Omron Sysmac Studio project TP - Automaçao (Sysmac Studio 1.56.0.64011, StandardProject)

# Controller new_Controller_0: NX1P2-9B24DT1 version 1.42
Task PrimaryTask (priority 4, period or condition 4000): Program0
Library OEN_Communication_V1_0_22 1.0.22 (contents left out)

VAR_GLOBAL
    Trama : ARRAY[0..3] OF OEN\Modbus\sModbusReq := [(Enable := True, NodeAdr := 1, FunctionCode := Fn02_ReadDiscreteInputs, Read := (StartAddressRemote := 0, StartAddressLocal := 0, Count := 49), Write := (StartAddressRemote := 0, StartAddressLocal := 0, Count := 0)), (Enable := True, NodeAdr := 1, FunctionCode := Fn15_WriteMultipleCoils, Read := (StartAddressRemote := 0, StartAddressLocal := 0, Count := 0), Write := (StartAddressRemote := 0, StartAddressLocal := 0, Count := 129)), (Enable := True, NodeAdr := 1, FunctionCode := Fn04_ReadInputRegisters, Read := (StartAddressRemote := 0, StartAddressLocal := 0, Count := 10), Write := (StartAddressRemote := 0, StartAddressLocal := 0, Count := 0)), (Enable := True, NodeAdr := 1, FunctionCode := Fn16_WriteMultipleRegisters, Read := (StartAddressRemote := 0, StartAddressLocal := 0, Count := 0), Write := (StartAddressRemote := 0, StartAddressLocal := 0, Count := 10))];  (* Trama *)
    out_Dig : ARRAY[0..130] OF BOOL;  (* Saidas digitais *)
    in_Dig : ARRAY[0..50] OF BOOL;  (* Entradas digitais *)
    in_Analog : ARRAY[0..10] OF WORD;  (* Entradas analogicas *)
    out_Analog : ARRAY[0..10] OF WORD;  (* Saidas analogicas *)
    BIO_Input_Bit_00 : BOOL;  (* Botão fisico; at BuiltInIO://cpu/#0/Input_Bit_00 *)
    BIO_Output_Bit_00 : BOOL;  (* Led Verde - Fisico; at BuiltInIO://cpu/#0/Output_Bit_00 *)
    BIO_Output_Bit_01 : BOOL;  (* Led Amarelo - Fisico; at BuiltInIO://cpu/#0/Output_Bit_01 *)
    BIO_Output_Bit_02 : BOOL;  (* Led Vermelho - Fisico; at BuiltInIO://cpu/#0/Output_Bit_02 *)
    ANALOG_Ch1_Analog_Output_Value : INT;  (* at BuiltInIO://opt/#0/Ch1_Analog_Output_Value *)
    Encomenda_Azul : DINT;  (* Numero de peça desta cor por encomenda *)
    Encomenda_Verde : DINT;  (* Numero de peça desta cor por encomenda *)
    Encomenda_Cinza : DINT;  (* Numero de peça desta cor por encomenda *)
    Peca_Boa_Azul : DINT;  (* Contador de peças boas produzidas *)
    Peca_Boa_Verde : DINT;  (* Contador de peças boas produzidas *)
    Peca_Boa_Cinza : DINT;  (* Contador de peças boas produzidas *)
    Peca_Lixo_Azul : DINT;  (* Contador de peças com defeito produzidas *)
    Peca_Lixo_Verde : DINT;  (* Contador de peças com defeito produzidas *)
    Peca_Lixo_Cinza : DINT;  (* Contador de peças com defeito produzidas *)
    Peca_Stock_Azul : DINT;  (* Contador de peças que foram para stock *)
    Peca_Stock_Verde : DINT;  (* Contador de peças que foram para stock *)
    Peca_Stock_Cinza : DINT;  (* Contador de peças que foram para stock *)
    HMI_Emitter : BOOL;
    HMI_R8 : BOOL;
    HMI_R0 : BOOL;
    HMI_R1 : BOOL;
    HMI_R3 : BOOL;
    HMI_R2 : BOOL;
    HMI_R4 : BOOL;
    HMI_R5 : BOOL;
    HMI_Alarme : BOOL;
    HMI_LG_10 : BOOL;
    HMI_LG_11 : BOOL;
    HMI_LG_12 : BOOL;
    HMI_LG_13 : BOOL;
    HMI_LG_14 : BOOL;
    HMI_LG_15 : BOOL;
    HMI_LG_18 : BOOL;
    HMI_LG_19 : BOOL;
    HMI_LY_10 : BOOL;
    HMI_LY_11 : BOOL;
    HMI_LY_12 : BOOL;
    HMI_LY_13 : BOOL;
    HMI_LY_14 : BOOL;
    HMI_LY_15 : BOOL;
    HMI_LY_18 : BOOL;
    HMI_LY_19 : BOOL;
    HMI_LR_10 : BOOL;
    HMI_LR_11 : BOOL;
    HMI_LR_12 : BOOL;
    HMI_LR_13 : BOOL;
    HMI_LR_14 : BOOL;
    HMI_LR_15 : BOOL;
    HMI_LR_18 : BOOL;
    HMI_LR_19 : BOOL;
    HMI_PP0_X : BOOL;
    HMI_PP1_X : BOOL;
    HMI_PP2_X : BOOL;
    HMI_PP0_Z : BOOL;
    HMI_PP1_Z : BOOL;
    HMI_PP2_Z : BOOL;
    HMI_PP0_Grab : BOOL;
    HMI_PP1_Grab : BOOL;
    HMI_PP2_Grab : BOOL;
    HMI_PP0_CW : BOOL;
    HMI_PP1_CW : BOOL;
    HMI_PP2_CW : BOOL;
    HMI_PP0_CCW : BOOL;
    HMI_PP1_CCW : BOOL;
    HMI_PP2_CCW : BOOL;
    HMI_DS0 : BOOL;
    HMI_DS1 : BOOL;
    HMI_DS2 : BOOL;
    HMI_DS3 : BOOL;
    HMI_DS4 : BOOL;
    HMI_DS5 : BOOL;
    HMI_DS6 : BOOL;
    HMI_DS7 : BOOL;
    HMI_DS8 : BOOL;
    HMI_DS9 : BOOL;
    HMI_DS10 : BOOL;
    HMI_DS11 : BOOL;
    HMI_DS12 : BOOL;
    HMI_DS13 : BOOL;
    HMI_DS14 : BOOL;
    HMI_DS15 : BOOL;
    HMI_DS16 : BOOL;
    HMI_DS17 : BOOL;
    HMI_DS18 : BOOL;
    HMI_DS19 : BOOL;
    HMI_DS20 : BOOL;
    HMI_DS21 : BOOL;
    HMI_DS22 : BOOL;
    HMI_DS23 : BOOL;
    HMI_DS24 : BOOL;
    HMI_DS25 : BOOL;
    HMI_DS26 : BOOL;
    HMI_DS27 : BOOL;
    HMI_DS28 : BOOL;
    HMI_T20 : BOOL;
    HMI_T21 : BOOL;
    HMI_T22 : BOOL;
    HMI_T23 : BOOL;
    HMI_T24 : BOOL;
    HMI_T25 : BOOL;
    HMI_T26 : BOOL;
    HMI_T27 : BOOL;
    HMI_T28 : BOOL;
    HMI_T29 : BOOL;
    HMI_T210 : BOOL;
    HMI_T211 : BOOL;
    HMI_T212 : BOOL;
    HMI_T213 : BOOL;
    HMI_T214 : BOOL;
    HMI_T215 : BOOL;
    HMI_T216 : BOOL;
    HMI_T217 : BOOL;
    HMI_T218 : BOOL;
    HMI_T219 : BOOL;
    HMI_T220 : BOOL;
    HMI_T221 : BOOL;
    HMI_T222 : BOOL;
    HMI_T223 : BOOL;
    HMI_T224 : BOOL;
    HMI_T225 : BOOL;
    HMI_T226 : BOOL;
    HMI_T227 : BOOL;
    HMI_T229 : BOOL;
    HMI_T230 : BOOL;
    HMI_T40 : BOOL;
    HMI_T41 : BOOL;
    HMI_T42 : BOOL;
    HMI_T43 : BOOL;
    HMI_T45 : BOOL;
    HMI_T46 : BOOL;
    HMI_T60 : BOOL;
    HMI_T61 : BOOL;
    HMI_T62 : BOOL;
    HMI_T63 : BOOL;
    HMI_T64 : BOOL;
    HMI_T65 : BOOL;
    HMI_T66 : BOOL;
    HMI_T67 : BOOL;
    HMI_T68 : BOOL;
    HMI_T69 : BOOL;
    HMI_CCW1 : BOOL;
    HMI_CCW0 : BOOL;
    HMI_CW2 : BOOL;
    HMI_CW3 : BOOL;
    HMI_CW4 : BOOL;
    HMI_CW5 : BOOL;
    HMI_CCW6 : BOOL;
    HMI_CCW7 : BOOL;
    HMI_CW8 : BOOL;
    HMI_CW9 : BOOL;
    HMI_CW10 : BOOL;
    HMI_CW11 : BOOL;
    HMI_CW12 : BOOL;
    HMI_CCW14 : BOOL;
    HMI_CW15 : BOOL;
    HMI_CW16 : BOOL;
    HMI_CW17 : BOOL;
    HMI_CW18 : BOOL;
    HMI_CCW20 : BOOL;
    HMI_CW21 : BOOL;
    HMI_PA3_Turn : BOOL;
    HMI_PA4_Turn : BOOL;
    HMI_PA3_Power : BOOL;
    HMI_PA4_Power : BOOL;
    HMI_B0_Power : BOOL;
    HMI_B1_Power : BOOL;
    HMI_B2_Power : BOOL;
    HMI_L0 : BOOL;
    HMI_L1 : BOOL;
    HMI_L2 : BOOL;
    HMI_MCS_0 : BOOL;
    HMI_MCS_1 : BOOL;
    HMI_MCS_2 : BOOL;
    Terminar_sessao : BOOL;  (* Sai do modo de manutenção da HMI *)
    HMI_Emissor : BOOL;
    HMI_Led_producao : BOOL;
    HMI_Led_Manutencao : BOOL;
    HMI_PP3_CCW : BOOL;
    HMI_PP3_CW : BOOL;
    HMI_BT_Linha_Principal : BOOL;
    HMI_BT_Linha_Azul : BOOL;
    HMI_BT_Linha_Verde : BOOL;
    HMI_BT_Linha_Cinza : BOOL;
    HMI_BT_Linha_Recolha : BOOL;
    VS : DINT;  (* Vision sensor *)
    Flag_Stop : BOOL;
    DS16 : BOOL;
    Encomenda_Total : DINT;
    DS28 : BOOL;
    BTSL_1 : BOOL;  (* Botão Seletor - posição 1 *)
    Page_Access : BOOL;
    HMI_Encomenda_Azul_Historico : ARRAY[1..10] OF REAL;
    HMI_Encomenda_Verde_Historico : ARRAY[1..10] OF REAL;
    HMI_Encomenda_Cinza_Historico : ARRAY[1..10] OF REAL;
    HMI_Historico_Index : INT := 1;
    Page_Access1 : BOOL;
    HMI_VoltaP : BOOL;
    HMI_VoltaRC : BOOL;
    HMI_Volta1 : BOOL;
    HMI_Volta2 : BOOL;
    HMI_Volta3 : BOOL;
    Encomenda_Pronta : BOOL;
    HMI_Flag_Stop : BOOL;
    HMI_VS : DINT;
    HMI_DS29 : BOOL;
    HMI_DS30 : BOOL;
    HMI_DS31 : BOOL;
    HMI_DS33 : BOOL;
    HMI_DS34 : BOOL;
    HMI_DS32 : BOOL;
    HMI_Emergencia : BOOL;
END_VAR

PROGRAM Program0
VAR
    ModBus_Client_PLC : OEN\Modbus\ModbusTCP_Client;  (* Bloco ModBus *)
    L0 : BOOL;  (* Lamina stop 0 *)
    L1 : BOOL;  (* Lamina stop 1 *)
    L2 : BOOL;  (* Lamina stop 2 *)
    Emitter : BOOL;  (* Emissor de peças *)
    R0 : BOOL;  (* Peças para o lixo *)
    R1 : BOOL;  (* Peças para o lixo *)
    R2 : BOOL;  (* Peças para stock *)
    R3 : BOOL;  (* Peças para o lixo *)
    R4 : BOOL;  (* Peças para stock *)
    R5 : BOOL;  (* Peças para stock *)
    R8 : BOOL;  (* Remove encomenda final *)
    BTSL_0 : BOOL;  (* Botão Seletor - posição 0 *)
    BTS : BOOL;  (* Botão Start *)
    BTE : BOOL;  (* Botão Emergencia *)
    BTSP : BOOL;  (* Botão Stop *)
    BTR : BOOL;  (* Botão Reset *)
    A2 : BOOL;  (* Alarme *)
    LG_10 : BOOL;  (* Led Verde - semaforo 10 *)
    LG_11 : BOOL;  (* Led Verde - semaforo 11 *)
    LG_12 : BOOL;  (* Led Verde - semaforo 12 *)
    LG_13 : BOOL;  (* Led Verde - semaforo 13 *)
    LG_14 : BOOL;  (* Led Verde - semaforo 14 *)
    LG_15 : BOOL;  (* Led Verde - semaforo 15 *)
    LG_18 : BOOL;  (* Led Verde - semaforo 18 *)
    LG_19 : BOOL;  (* Led Verde - semaforo 19 *)
    LR_10 : BOOL;  (* Led Vermelho - semaforo 10 *)
    LR_11 : BOOL;  (* Led Vermelho - semaforo 11 *)
    LR_12 : BOOL;  (* Led Vermelho - semaforo 12 *)
    LR_13 : BOOL;  (* Led Vermelho - semaforo 13 *)
    LR_14 : BOOL;  (* Led Vermelho - semaforo 14 *)
    LR_15 : BOOL;  (* Led Vermelho - semaforo 15 *)
    LR_18 : BOOL;  (* Led Vermelho - semaforo 18 *)
    LR_19 : BOOL;  (* Led Vermelho - semaforo 19 *)
    LY_10 : BOOL;  (* Led Amarelo - semaforo 10 *)
    LY_11 : BOOL;  (* Led Amarelo - semaforo 11 *)
    LY_12 : BOOL;  (* Led Amarelo - semaforo 12 *)
    LY_13 : BOOL;  (* Led Amarelo - semaforo 13 *)
    LY_14 : BOOL;  (* Led Amarelo - semaforo 14 *)
    LY_15 : BOOL;  (* Led Amarelo - semaforo 15 *)
    LY_18 : BOOL;  (* Led Amarelo - semaforo 18 *)
    LY_19 : BOOL;  (* Led Amarelo - semaforo 19 *)
    DS0 : BOOL;  (* Opto-Switch 0 *)
    DS1 : BOOL;  (* Opto-Switch 1 *)
    DS2 : BOOL;  (* Opto-Switch 2 *)
    DS3 : BOOL;  (* Opto-Switch 3 *)
    DS4 : BOOL;  (* Opto-Switch 4 *)
    DS5 : BOOL;  (* Opto-Switch 5 *)
    DS6 : BOOL;  (* Opto-Switch 6 *)
    DS7 : BOOL;  (* Opto-Switch 7 *)
    DS8 : BOOL;  (* Opto-Switch 8 *)
    DS9 : BOOL;  (* Opto-Switch 9 *)
    DS10 : BOOL;  (* Opto-Switch 10 *)
    DS11 : BOOL;  (* Opto-Switch 11 *)
    DS12 : BOOL;  (* Opto-Switch 12 *)
    DS13 : BOOL;  (* Opto-Switch 13 *)
    DS14 : BOOL;  (* Opto-Switch 14 *)
    DS15 : BOOL;  (* Opto-Switch 15 *)
    DS16 : BOOL;  (* Opto-Switch 16 *)
    DS29 : BOOL;  (* Opto-Switch 29 *)
    DS30 : BOOL;  (* Opto-Switch 30 *)
    DS31 : BOOL;  (* Opto-Switch 31 *)
    DS32 : BOOL;  (* Opto-Switch 32 *)
    DS33 : BOOL;  (* Opto-Switch 33 *)
    DS34 : BOOL;  (* Opto-Switch 34 *)
    DS17 : BOOL;  (* Opto-Switch 17 *)
    DS18 : BOOL;  (* Opto-Switch 18 *)
    DS19 : BOOL;  (* Opto-Switch 19 *)
    DS20 : BOOL;  (* Opto-Switch 20 *)
    DS21 : BOOL;  (* Opto-Switch 21 *)
    DS22 : BOOL;  (* Opto-Switch 22 *)
    DS23 : BOOL;  (* Opto-Switch 23 *)
    DS24 : BOOL;  (* Opto-Switch 24 *)
    DS25 : BOOL;  (* Opto-Switch 25 *)
    DS26 : BOOL;  (* Opto-Switch 26 *)
    DS27 : BOOL;  (* Opto-Switch 27 *)
    DS28 : BOOL;  (* Opto-Switch 28 *)
    PP0_Detect : BOOL;  (* Sensor que dedeta peça na Pick and Place 0 *)
    PP1_Detect : BOOL;  (* Sensor que dedeta peça na Pick and Place 1 *)
    PP2_Detect : BOOL;  (* Sensor que dedeta peça na Pick and Place 2 *)
    PP0_X : BOOL;  (* Pick and place 0 - eixo x *)
    PP1_X : BOOL;  (* Pick and place 1 - eixo x *)
    PP2_X : BOOL;  (* Pick and place 2 - eixo x *)
    PP0_Z : BOOL;  (* Pick and place 0 - eixo z *)
    PP1_Z : BOOL;  (* Pick and place 1 - eixo z *)
    PP2_Z : BOOL;  (* Pick and place 2 - eixo z *)
    PP0_Grab : BOOL;  (* Pick and place 0 - agarra peça *)
    PP1_Grab : BOOL;  (* Pick and place 1 - agarra peça *)
    PP2_Grab : BOOL;  (* Pick and place 2 - agarra peça *)
    PP0_CW : BOOL;  (* Pick and place 0 - roda no sentido horario *)
    PP1_CW : BOOL;  (* Pick and place 1 - roda no sentido horario *)
    PP2_CW : BOOL;  (* Pick and place 2 - roda no sentido horario *)
    PP0_CCW : BOOL;  (* Pick and place 0 - roda no sentido anti horario *)
    PP1_CCW : BOOL;  (* Pick and place 1 - roda no sentido anti horario *)
    PP2_CCW : BOOL;  (* Pick and place 2 - roda no sentido anti horario *)
    CCW0 : BOOL;  (* Tapete curvo 0 *)
    CCW1 : BOOL;  (* Tapete curvo 1 *)
    CW2 : BOOL;  (* Tapete curvo 2 *)
    CW3 : BOOL;  (* Tapete curvo 3 *)
    CW4 : BOOL;  (* Tapete curvo 4 *)
    CW5 : BOOL;  (* Tapete curvo 5 *)
    CCW6 : BOOL;  (* Tapete curvo 6 *)
    CCW7 : BOOL;  (* Tapete curvo 7 *)
    CW8 : BOOL;  (* Tapete curvo 8 *)
    CW9 : BOOL;  (* Tapete curvo 9 *)
    CW10 : BOOL;  (* Tapete curvo 10 *)
    CW11 : BOOL;  (* Tapete curvo 11 *)
    CW12 : BOOL;  (* Tapete curvo 12 *)
    CCW14 : BOOL;  (* Tapete curvo 14 *)
    CW15 : BOOL;  (* Tapete curvo 15 *)
    CW16 : BOOL;  (* Tapete curvo 16 *)
    CW17 : BOOL;  (* Tapete curvo 17 *)
    CW18 : BOOL;  (* Tapete curvo 18 *)
    CCW20 : BOOL;  (* Tapete curvo 20 *)
    CW21 : BOOL;  (* Tapete curvo 21 *)
    T20 : BOOL;  (* Tapete 2m n0 *)
    T21 : BOOL;  (* Tapete 2m n1 *)
    T22 : BOOL;  (* Tapete 2m n2 *)
    T23 : BOOL;  (* Tapete 2m n3 *)
    T24 : BOOL;  (* Tapete 2m n4 *)
    T25 : BOOL;  (* Tapete 2m n5 *)
    T26 : BOOL;  (* Tapete 2m n6 *)
    T27 : BOOL;  (* Tapete 2m n7 *)
    T28 : BOOL;  (* Tapete 2m n8 *)
    T29 : BOOL;  (* Tapete 2m n9 *)
    T210 : BOOL;  (* Tapete 2m n10 *)
    T211 : BOOL;  (* Tapete 2m n11 *)
    T212 : BOOL;  (* Tapete 2m n12 *)
    T213 : BOOL;  (* Tapete 2m n13 *)
    T214 : BOOL;  (* Tapete 2m n14 *)
    T215 : BOOL;  (* Tapete 2m n15 *)
    T216 : BOOL;  (* Tapete 2m n16 *)
    T217 : BOOL;  (* Tapete 2m n17 *)
    T218 : BOOL;  (* Tapete 2m n18 *)
    T219 : BOOL;  (* Tapete 2m n19 *)
    T220 : BOOL;  (* Tapete 2m n20 *)
    T221 : BOOL;  (* Tapete 2m n21 *)
    T222 : BOOL;  (* Tapete 2m n22 *)
    T223 : BOOL;  (* Tapete 2m n23 *)
    T224 : BOOL;  (* Tapete 2m n24 *)
    T225 : BOOL;  (* Tapete 2m n25 *)
    T226 : BOOL;  (* Tapete 2m n26 *)
    T227 : BOOL;  (* Tapete 2m n27 *)
    T229 : BOOL;  (* Tapete 2m n29 *)
    T230 : BOOL;  (* Tapete 2m n30 *)
    T40 : BOOL;  (* Tapete 4m n0 *)
    T41 : BOOL;  (* Tapete 4m n1 *)
    T42 : BOOL;  (* Tapete 4m n2 *)
    T43 : BOOL;  (* Tapete 4m n3 *)
    T45 : BOOL;  (* Tapete 4m n5 *)
    T46 : BOOL;  (* Tapete 4m n6 *)
    T60 : BOOL;  (* Tapete 6m n0 *)
    T61 : BOOL;  (* Tapete 6m n1 *)
    T62 : BOOL;  (* Tapete 6m n2 *)
    T63 : BOOL;  (* Tapete 6m n3 *)
    T64 : BOOL;  (* Tapete 6m n4 *)
    T65 : BOOL;  (* Tapete 6m n5 *)
    T66 : BOOL;  (* Tapete 6m n6 *)
    T67 : BOOL;  (* Tapete 6m n7 *)
    T68 : BOOL;  (* Tapete 6m n8 *)
    T69 : BOOL;  (* Tapete 6m n9 *)
    B0_W : INT;  (* Balança 0 - peso *)
    B1_W : INT;  (* Balança 1 - peso *)
    B2_W : INT;  (* Balança 2 - peso *)
    B0_Power : BOOL;  (* Balança 0 - tapete anda para a frente *)
    B1_Power : BOOL;  (* Balança 1 - tapete anda para a frente *)
    B2_Power : BOOL;  (* Balança 2 - tapete anda para a frente *)
    PA3_Power : BOOL;  (* Pivot Arm 3 - tapete anda para a frente *)
    PA3_Turn : BOOL;  (* Pivot Arm 3 - rodar *)
    PA4_Power : BOOL;  (* Pivot Arm 4 - tapete anda para a frente *)
    PA4_Turn : BOOL;  (* Pivot Arm 4 - rotação *)
    MCS_0 : BOOL;  (* Machine Center 0 - start *)
    MCS_1 : BOOL;  (* Machine Center 1 - start *)
    MCS_2 : BOOL;  (* Machine Center 2 - start *)
    Arranque : INT;  (* Etapas do arranque da linha completa *)
    Tapete_Princioal : INT;  (* Etapas que controlam o inicio da produção *)
    Inicio_Linha_A : INT;  (* Etapa para controlar 1º tapete da linha *)
    Inicio_Linha_V : INT;  (* Etapa para controlar 1º tapete da linha *)
    Inicio_Linha_C : INT;  (* Etapa para controlar 1º tapete da linha *)
    PintaSeca_Azul : INT;  (* Etapas para pintar e secar a peça Azul *)
    PintaSeca_Verde : INT;  (* Etapas para pintar e secar a peça Verde *)
    PintaSeca_Cinza : INT;  (* Etapas para pintar e secar a peça Cinza *)
    Balaca_A : INT;  (* Etapas que controlam o tapete da balaça *)
    Balaca_V : INT;  (* Etapas que controlam o tapete da balaça *)
    Balaca_C : INT;  (* Etapas que controlam o tapete da balaça *)
    Analisa_Azul : INT;  (* Etapas para decidir o que faz com a peça a partir do peso *)
    Analisa_Verde : INT;  (* Etapas para decidir o que faz com a peça a partir do peso *)
    Analisa_Cinza : INT;  (* Etapas para decidir o que faz com a peça a partir do peso *)
    Boa_Azul : INT;  (* Etapas para as peças boas *)
    Boa_Verde : INT;  (* Etapas para as peças boas *)
    Boa_Cinza : INT;  (* Etapas para as peças boas *)
    ParaReparar_Azul : INT;  (* Etapas para quando a peça azul tem que ser reparada *)
    ParaReparar_Verde : INT;  (* Etapas para quando a peça verde tem que ser reparada *)
    ParaReparar_Cinza : INT;  (* Etapas para quando a peça cinza tem que ser reparada *)
    Stock_Azul : INT;  (* Etapas para quando a encomenda já tem o maximo de peças de uma encomenda *)
    Stock_Verde : INT;  (* Etapas para quando a encomenda já tem o maximo de peças de uma encomenda *)
    Stock_Cinza : INT;  (* Etapas para quando a encomenda já tem o maximo de peças de uma encomenda *)
    Lixo_Azul : INT;  (* Etapas para quando a peça azul é defeituosa *)
    Lixo_Verde : INT;  (* Etapas para quando a peça verde é defeituosa *)
    Lixo_Cinza : INT;  (* Etapas para quando a peça cinza é defeituosa *)
    Recolhe_Boa_Azul : INT;  (* Etapas para levar as peças boas até ao local comum de recolha *)
    Recolhe_Boa_Verde : INT;  (* Etapas para levar as peças boas até ao local comum de recolha *)
    Recolhe_Boa_Cinza : INT;  (* Etapas para levar as peças boas até ao local comum de recolha *)
    Recolha_Comum : INT;  (* Etapas para a recolha comum das peças até à palete *)
END_VAR
VAR CONSTANT
    VSA_B : INT := 3;  (* Peça azul - boa *)
    VSV_B : INT := 6;  (* Peça verde - boa *)
    VSC_B : INT := 9;  (* Peça cinza - boa *)
    VSA_PR : INT := 1;  (* Peça azul - para reparar *)
    VSV_PR : INT := 4;  (* Peça verde - para reparar *)
    VSC_PR : INT := 7;  (* Peça cinza - para reparar *)
    VSA_L : INT := 2;  (* Peça azul - lixo *)
    VSV_L : INT := 5;  (* Peça verde - lixo *)
    VSC_L : INT := 8;  (* Peça cinza - lixo *)
END_VAR
VAR
    BC_Peso : REAL;  (* Peso atual da peça - cinza *)
    BA_Peso : REAL;  (* Peso atual da peça - azul *)
    BV_Peso : REAL;  (* Peso atual da peça - verde *)
    Manutencao_LP : INT;  (* Etapas para a anutenção da linha principal *)
    Manutencao_LA : INT;  (* Etapas para a anutenção da linha azul *)
    Manutencao_LV : INT;  (* Etapas para a anutenção da linha verde *)
    Manutencao_LC : INT;  (* Etapas para a anutenção da linha cinza *)
    Manutencao_LR : INT;  (* Etapas para a anutenção da linha de recolha *)
    Flag_BusyPP1 : BOOL;  (* Flag que indica se a pick and place está a ser usada *)
    VS : INT;  (* Vision Sensor *)
    Flag_Stop : BOOL;  (* Flag para ativar modo de STOP *)
    Flag_ModoProd : BOOL;  (* Flag para ativar etapas do modo de produção *)
    Flag_Inicio_Linha_Azul : BOOL;  (* Flag para iniciar a linha azul *)
    Flag_Inicio_Linha_Verde : BOOL;  (* Flag para iniciar a linha verde *)
    Flag_Inicio_Linha_Cinza : BOOL;  (* Flag para iniciar a linha azul *)
    Flag_PintaSeca_A : BOOL;  (* Flag para iniciar as etapas de pintura e secagem da peça *)
    Flag_Pesagem_A : BOOL;  (* Etapas para a zona de pesagem *)
    Flag_Balaca_A : BOOL;  (* Flag para andar balaça da peça *)
    Flag_Analisa_A : BOOL;  (* Flag para analisar peso da peça *)
    Flag_Boa_A : BOOL;  (* Flag para ativar etapas se a peça AZUL é boa *)
    Flag_ParaReparar_A : BOOL;  (* Flag para ativar etapas se a peça AZUL é para reparar *)
    Flag_Lixo_A : BOOL;  (* Flag para ativar etapas se a peça AZUL é lixo *)
    Flag_Stock_A : BOOL;  (* Flag para ativar etapas se a peça AZUL é para stock *)
    Flag_Analisa_C : BOOL;  (* Flag para analisar peso da peça *)
    Flag_Analisa_V : BOOL;  (* Flag para analisar peso da peça *)
    Flag_Boa_V : BOOL;  (* Flag para ativar etapas se a peça VERDE é boa *)
    Flag_ParaReparar_V : BOOL;  (* Flag para ativar etapas se a peça VERDE é para reparar *)
    Flag_Lixo_V : BOOL;  (* Flag para ativar etapas se a peça VERDE é lixo *)
    Flag_Stock_V : BOOL;  (* Flag para ativar etapas se a peça VERDE é para stock *)
    Flag_Boa_C : BOOL;  (* Flag para ativar etapas se a peça CINZA é boa *)
    Flag_ParaReparar_C : BOOL;  (* Flag para ativar etapas se a peça CINZA é para reparar *)
    Flag_Lixo_C : BOOL;  (* Flag para ativar etapas se a peça CINZA é lixo *)
    Flag_Stock_C : BOOL;  (* Flag para ativar etapas se a peça CINZA é para stock *)
    Flag_RecolheBoa_A : BOOL;  (* Flag para ativar etapas para levar a peça até zona de recolha comum *)
    Entra_Boa_Azul : INT := 0;  (* Conta que entrou uma peça BOA para a zona de recolha *)
    Sai_Azul : INT;
    Flag_RecolhaComum : BOOL;  (* Flag que ativa a zona de recolha comum *)
    Flag_Reset_Boas_A : BOOL;
    Encomenda_V : INT;  (* Nº de peças VERDES necessárias para competar a encomenda *)
    Encomenda_C : INT;  (* Nº de peças CINZAS necessárias para competar a encomenda *)
    Encomenda_A : INT;  (* Nº de peças AZUIS necessárias para competar a encomenda *)
    Encomenda_T : INT;  (* Nº de encomendas completadas *)
    ContadorPecasBoasAzuis : CTU;
    ContadorPecasBoasVerdes : CTU;
    ContadorPecasBoasCinzas : CTU;
    Conta_Pecas_Boas_A : INT;  (* Contador de peças boas produzidas até terminar encomenda. *)
    Conta_Pecas_Boas_V : INT;  (* Contador de peças boas produzidas até terminar encomenda. *)
    Conta_Pecas_Boas_C : INT;  (* Contador de peças boas produzidas até terminar encomenda. *)
    Conta_Pecas_Lixo_A : INT;  (* Contador de peças com defeito produzidas até terminar encomenda. *)
    Conta_Pecas_Lixo_V : INT;  (* Contador de peças com defeito produzidas até terminar encomenda. *)
    Conta_Pecas_Lixo_C : INT;  (* Contador de peças com defeito produzidas até terminar encomenda. *)
    Conta_Pecas_Stock_A : INT;  (* Contador de peças para stock *)
    Conta_Pecas_Stock_V : INT;  (* Contador de peças para stock *)
    Conta_Pecas_Stock_C : INT;  (* Contador de peças para stock *)
    ContadorPecasStockAzuis : CTU;
    Flag_Reset_Boas_V : BOOL;
    ContadorPecasStockVerdes : CTU;
    Flag_Reset_Boas_C : BOOL;
    ContadorPecasStockCinzas : CTU;
    ContaEntradaBoaAzul : CTU;
    ContaSaidaAzul : CTU;
    Passou_1s_A1 : BOOL;
    Flag_RecolheLixo_A : BOOL;
    Timer1_Azul : TON;
    Recolhe_Lixo_Azul : INT;  (* Etapas que levam a peça até ao lixo *)
    ContaEntradaVerde : CTU;
    ContaSaidaVerde : CTU;
    ContaEntradaCinza : CTU;
    ContaSaidaCinza : CTU;
    Entra_Boa_Verde : INT := 0;  (* Conta que entrou uma peça BOA para a zona de recolha *)
    Entra_Boa_Cinza : INT := 0;  (* Conta que entrou uma peça BOA para a zona de recolha *)
    Recolhe_Lixo_Verde : INT;  (* Etapas que levam a peça até ao lixo *)
    Recolhe_Lixo_Cinza : INT;  (* Etapas que levam a peça até ao lixo *)
    Flag_Balaca_V : BOOL;  (* Flag para andar balaça da peça *)
    Flag_Balaca_C : BOOL;  (* Flag para andar balaça da peça *)
    Flag_BusyPP2 : BOOL;  (* Flag que indica se a pick and place está a ser usada *)
    Flag_BusyPP0 : BOOL;  (* Flag que indica se a pick and place está a ser usada *)
    Flag_Pesagem_V : BOOL;  (* Etapas para a zona de pesagem *)
    Flag_Pesagem_C : BOOL;  (* Etapas para a zona de pesagem *)
    Passou_1s_V1 : INT;
    Passou_1s_C1 : INT;
    Timer1_Verde : TON;
    Timer1_Cinza : TON;
    Sai_Verde : INT;
    Sai_Cinza : INT;
    Flag_RecolheBoa_V : BOOL;
    Flag_RecolheBoa_C : BOOL;
    Flag_PintaSeca_V : BOOL;  (* Flag para iniciar as etapas de pintura e secagem da peça *)
    Flag_PintaSeca_C : BOOL;  (* Flag para iniciar as etapas de pintura e secagem da peça *)
    Flag_RecolheLixo_V : BOOL;
    Flag_RecolheLixo_C : BOOL;
    Flag_Trasporta_Peca_Reparada_A : BOOL;
    Flag_Trasporta_Peca_Reparada_V : BOOL;
    Flag_Trasporta_Peca_Reparada_C : BOOL;
    Transporte_RP_A : INT;
    Transporte_RP_V : INT;
    Transporte_RP_C : INT;
    Flag_Sai_CNC_A : BOOL;
    Flag_Sai_CNC_V : BOOL;
    Flag_Sai_CNC_C : BOOL;
    Passou_3s_A : BOOL;
    Passou_3s_V : BOOL;
    Passou_3s_C : BOOL;
    Saida_CNC_A : INT;
    Saida_CNC_V : INT;
    Saida_CNC_C : INT;
    Timer2_Azul : TON;
    Passou_1s_A2 : BOOL;
    Timer3_Azul : TON;
    Flag_Transporte_Stock_A : BOOL;
    Recolhe_Stock_A : INT;
    Recolhe_Stock_V : INT;
    Recolhe_Stock_C : INT;
    Flag_Transporte_Stock_V : BOOL;
    Flag_Transporte_Stock_C : BOOL;
    Reset_Contadores : BOOL;
    ContaEntradaParaRepararAzul : CTU;
    Entra_PR_Azul : INT := 0;
    Entra_PR_Verde : INT;
    Entra_PR_Cinza : INT := 0;
    ContadorPecasLixoAzuis : CTU;
    ContadorPecasLixoVerdes : CTU;
    ContadorPecasLixoCinzas : CTU;
    ContadorPecasReparadasAzuis : CTU;
    Conta_Pecas_Reparadas_A : INT;  (* Conta peça reparada *)
    ContadorPecasReparadasVerdes : CTU;
    Conta_Pecas_Reparadas_V : INT;  (* Conta peça reparada *)
    ContadorPecasReparadasCinzas : CTU;
    Conta_Pecas_Reparadas_C : INT;  (* Conta peça reparada *)
    ContaTotal_Azul : INT;
    Diferenca_Azuis : INT;  (* Quantas peças boas ainda estão no tapete *)
    Passou_3s_A2 : BOOL;
    Timer4_Azul : TON;
    timer1_F : BOOL;  (* Timer acabou *)
    timer2_F : BOOL;  (* Timer acabou *)
    Timer1 : TON;
    Timer2 : TON;
    timer3_F : BOOL;  (* Timer acabou *)
    Timer3 : TON;
    timer4_F : BOOL;  (* Timer acabou *)
    Timer4 : TON;
    timer5_F : BOOL;  (* Timer acabou *)
    Timer5 : TON;
    timer6_F : BOOL;  (* Timer acabou *)
    timer7_F : BOOL;  (* Timer acabou *)
    timer8_F : BOOL;  (* Timer acabou *)
    timer9_F : BOOL;  (* Timer acabou *)
    Timer6 : TON;
    Timer7 : TON;
    Timer8 : TON;
    ContaSaida_A : INT;
    Timer9 : TON;
    timer10_F : BOOL;  (* Timer acabou *)
    Timer10 : TON;
    timer11_F : BOOL;  (* Timer acabou *)
    Timer11 : TON;
    timer12_F : BOOL;  (* Timer acabou *)
    Timer12 : TON;
    Timer13 : TON;
    timer13_F : BOOL;  (* Timer acabou *)
    timer14_F : BOOL;  (* Timer acabou *)
    Timer14 : TON;
    timer15_F : BOOL;  (* Timer acabou *)
    Timer15 : TON;
    timer16_F : BOOL;  (* Timer acabou *)
    Timer16 : TON;
    timer17_F : BOOL;  (* Timer acabou *)
    Timer17 : TON;
    timer18_F : BOOL;  (* Timer acabou *)
    Timer18 : TON;
    Timer19 : TON;
    timer19_F : BOOL;  (* Timer acabou *)
    timer20_F : BOOL;  (* Timer acabou *)
    timer21_F : BOOL;  (* Timer acabou *)
    Timer20 : TON;
    Timer21 : TON;
    cpla : BOOL;
    timer22_F : BOOL;  (* Timer acabou *)
    Timer22 : TON;
    timer23_F : BOOL;  (* Timer acabou *)
    Timer23 : TON;
    timer24_F : BOOL;  (* Timer acabou *)
    Timer24 : TON;
    timer25_F : BOOL;  (* Timer acabou *)
    Timer25 : TON;
    timer26_F : BOOL;  (* Timer acabou *)
    Timer26 : TON;
    timer27_F : BOOL;  (* Timer acabou *)
    Timer27 : TON;
    timer28_F : BOOL;  (* Timer acabou *)
    Timer28 : TON;
    ContadorPecasReparaAzuis : CTU;
    Conta_Peca_Boa_Reparadas_Azul : INT;  (* Peças reparadas e boas *)
    Flag_PP : BOOL;
    timer29_F : BOOL;  (* Timer acabou *)
    Timer29 : TON;
    timer30_F : BOOL;  (* Timer acabou *)
    Timer30 : TON;
    Conta_SaidaTapete : INT;  (* Conta quantas peças sairam do tapete da recolha comum *)
    ContaTotal : CTU;
    Total_Aux : INT;  (* Total auxiliar para saber o numero de peças da encomenda *)
    Total : INT;  (* Total de peças para a encomenda *)
    Timer31_F : BOOL;  (* Timer acabou *)
    Timer31 : TON;
    Timer32_F : BOOL;  (* Timer acabou *)
    Timer32 : TON;
    timer33_F : BOOL;  (* Timer acabou *)
    Timer34_F : BOOL;  (* Timer acabou *)
    Timer33 : TON;
    timer35_F : BOOL;  (* Timer acabou *)
    Timer34 : TON;
    Conta_Peca_Boa_Reparadas_Verde : INT;  (* Peças reparadas e boas *)
    Timer36_F : BOOL;  (* Timer acabou *)
    timer37_F : BOOL;  (* Timer acabou *)
    Timer35 : TON;
    Timer36 : TON;
    Timer37 : TON;
    Diferenca_Verde : INT;  (* Quantas peças boas ainda estão no tapete *)
    ContaSaida_V : INT;
    timer38_F : BOOL;  (* Timer acabou *)
    Timer38 : TON;
    Timer39_F : BOOL;  (* Timer acabou *)
    Timer39 : TON;
    timer40_F : BOOL;  (* Timer acabou *)
    timer41_F : BOOL;  (* Timer acabou *)
    timer42_F : BOOL;  (* Timer acabou *)
    timer43_F : BOOL;  (* Timer acabou *)
    timer44_F : BOOL;  (* Timer acabou *)
    Timer40 : TON;
    Timer41 : TON;
    Timer42 : TON;
    Timer43 : TON;
    Timer44 : TON;
    timer45_F : BOOL;  (* Timer acabou *)
    Timer45 : TON;
    timer46_F : BOOL;  (* Timer acabou *)
    timer47_F : BOOL;  (* Timer acabou *)
    timer48_F : BOOL;  (* Timer acabou *)
    timer49_F : BOOL;  (* Timer acabou *)
    timer50_F : BOOL;  (* Timer acabou *)
    timer51_F : BOOL;  (* Timer acabou *)
    Timer46 : TON;
    Timer47 : TON;
    Timer48 : TON;
    Timer49 : TON;
    Timer51 : TON;
    Timer50 : TON;
    timer52_F : BOOL;  (* Timer acabou *)
    Timer52 : TON;
    Timer53_F : BOOL;  (* Timer acabou *)
    timer54_F : BOOL;  (* Timer acabou *)
    Timer53 : TON;
    Timer54 : TON;
    timer55_F : BOOL;  (* Timer acabou *)
    timer56_F : BOOL;  (* Timer acabou *)
    timer57_F : BOOL;  (* Timer acabou *)
    timer58_F : BOOL;  (* Timer acabou *)
    timer59_F : BOOL;  (* Timer acabou *)
    timer60_F : BOOL;  (* Timer acabou *)
    timer61_F : BOOL;  (* Timer acabou *)
    timer62_F : BOOL;  (* Timer acabou *)
    timer63_F : BOOL;  (* Timer acabou *)
    Timer55 : TON;
    Timer56 : TON;
    Timer57 : TON;
    Timer58 : TON;
    Timer59 : TON;
    Timer60 : TON;
    Timer61 : TON;
    Timer62 : TON;
    Timer63 : TON;
    timer64_F : BOOL;  (* Timer acabou *)
    Timer64 : TON;
    Conta_Peca_Boa_Reparadas_CInza : INT;  (* Peças reparadas e boas *)
    Diferenca_Cinza : INT;  (* Quantas peças boas ainda estão no tapete *)
    ContaSaida_c : INT;
    timer65_F : BOOL;  (* Timer acabou *)
    Timer65 : TON;
    timer66_F : BOOL;  (* Timer acabou *)
    Timer67_F : BOOL;  (* Timer acabou *)
    Timer66 : TON;
    Timer67 : TON;
    timer68_F : BOOL;  (* Timer acabou *)
    Timer68 : TON;
    Timer69_F : BOOL;  (* Timer acabou *)
    timer70_F : BOOL;  (* Timer acabou *)
    Timer69 : TON;
    Timer70 : TON;
    timer71_F : BOOL;  (* Timer acabou *)
    Timer71 : TON;
    Timer72_F : BOOL;  (* Timer acabou *)
    Timer72 : TON;
    timer73_F : BOOL;  (* Timer acabou *)
    timer74_F : BOOL;  (* Timer acabou *)
    timer75_F : BOOL;  (* Timer acabou *)
    timer76_F : BOOL;  (* Timer acabou *)
    Timer73 : TON;
    Timer74 : TON;
    Timer75 : TON;
    Timer76 : TON;
    timer77_F : BOOL;  (* Timer acabou *)
    Timer77 : TON;
    timer78_F : BOOL;  (* Timer acabou *)
    Timer78 : TON;
    timer79_F : BOOL;  (* Timer acabou *)
    timer80_F : BOOL;  (* Timer acabou *)
    timer81_F : BOOL;  (* Timer acabou *)
    timer82_F : BOOL;  (* Timer acabou *)
    timer83_F : BOOL;  (* Timer acabou *)
    timer84_F : BOOL;  (* Timer acabou *)
    Timer79 : TON;
    Timer80 : TON;
    Timer81 : TON;
    Timer82 : TON;
    Timer83 : TON;
    Timer84 : TON;
    timer85_F : BOOL;  (* Timer acabou *)
    Timer85 : TON;
    Timer86_F : BOOL;  (* Timer acabou *)
    timer87_F : BOOL;  (* Timer acabou *)
    Timer86 : TON;
    Timer87 : TON;
    timer88_F : BOOL;  (* Timer acabou *)
    timer89_F : BOOL;  (* Timer acabou *)
    timer90_F : BOOL;  (* Timer acabou *)
    timer91_F : BOOL;  (* Timer acabou *)
    timer92_F : BOOL;  (* Timer acabou *)
    timer93_F : BOOL;  (* Timer acabou *)
    timer94_F : BOOL;  (* Timer acabou *)
    timer95_F : BOOL;  (* Timer acabou *)
    timer96_F : BOOL;  (* Timer acabou *)
    Timer88 : TON;
    Timer89 : TON;
    Timer90 : TON;
    Timer91 : TON;
    Timer92 : TON;
    Timer93 : TON;
    Timer94 : TON;
    Timer96 : TON;
    Timer95 : TON;
    timer97_F : BOOL;  (* Timer acabou *)
    Timer97 : TON;
    Timer100_F : BOOL;  (* Timer acabou *)
    Timer100 : TON;
    Timer101 : TON;
    timer101_F : BOOL;  (* Timer acabou *)
    Timer102 : TON;
    Timer102_F : BOOL;  (* Timer acabou *)
    Timer103 : TON;
    timer103_F : BOOL;  (* Timer acabou *)
    Timer104 : TON;
    timer104_F : BOOL;  (* Timer acabou *)
    Timer105 : TON;
    timer105_F : BOOL;  (* Timer acabou *)
    Timer106 : TON;
    Timer107 : TON;
    Timer108 : TON;
    Timer109 : TON;
    Timer110 : TON;
    Timer111 : TON;
    Timer112 : TON;
    Timer113 : TON;
    Timer114 : TON;
    Timer115 : TON;
    Timer116 : TON;
    Timer117 : TON;
    Timer118 : TON;
    Timer119 : TON;
    Timer120 : TON;
    Timer121 : TON;
    Timer122 : TON;
    Timer123 : TON;
    Timer124 : TON;
    Timer125 : TON;
    Timer126 : TON;
    Timer127 : TON;
    Timer128 : TON;
    Timer129 : TON;
    Timer130 : TON;
    Timer131 : TON;
    timer106_F : BOOL;  (* Timer acabou *)
    timer107_F : BOOL;  (* Timer acabou *)
    timer108_F : BOOL;  (* Timer acabou *)
    timer109_F : BOOL;  (* Timer acabou *)
    timer110_F : BOOL;  (* Timer acabou *)
    timer111_F : BOOL;  (* Timer acabou *)
    timer112_F : BOOL;  (* Timer acabou *)
    timer113_F : BOOL;  (* Timer acabou *)
    timer114_F : BOOL;  (* Timer acabou *)
    timer115_F : BOOL;  (* Timer acabou *)
    timer116_F : BOOL;  (* Timer acabou *)
    timer117_F : BOOL;  (* Timer acabou *)
    timer118_F : BOOL;  (* Timer acabou *)
    timer119_F : BOOL;  (* Timer acabou *)
    timer120_F : BOOL;  (* Timer acabou *)
    Timer121_F : BOOL;  (* Timer acabou *)
    timer122_F : BOOL;  (* Timer acabou *)
    timer123_F : BOOL;  (* Timer acabou *)
    timer124_F : BOOL;  (* Timer acabou *)
    timer125_F : BOOL;  (* Timer acabou *)
    timer126_F : BOOL;  (* Timer acabou *)
    timer127_F : BOOL;  (* Timer acabou *)
    timer128_F : BOOL;  (* Timer acabou *)
    timer129_F : BOOL;  (* Timer acabou *)
    timer130_F : BOOL;  (* Timer acabou *)
    timer131_F : BOOL;  (* Timer acabou *)
    Timer200 : TON;
    Timer201 : TON;
    Timer202 : TON;
    Timer203 : TON;
    Timer204 : TON;
    Timer205 : TON;
    Timer206 : TON;
    Timer207 : TON;
    Timer208 : TON;
    Timer209 : TON;
    Timer210 : TON;
    Timer211 : TON;
    Timer212 : TON;
    Timer213 : TON;
    Timer214 : TON;
    Timer215 : TON;
    Timer216 : TON;
    Timer217 : TON;
    Timer218 : TON;
    Timer219 : TON;
    Timer220 : TON;
    Timer221 : TON;
    Timer222 : TON;
    Timer223 : TON;
    Timer224 : TON;
    Timer225 : TON;
    Timer226 : TON;
    Timer227 : TON;
    Timer228 : TON;
    Timer229 : TON;
    Timer230 : TON;
    Timer231 : TON;
    Timer200_F : BOOL;  (* Timer acabou *)
    timer201_F : BOOL;  (* Timer acabou *)
    Timer202_F : BOOL;  (* Timer acabou *)
    timer203_F : BOOL;  (* Timer acabou *)
    timer204_F : BOOL;  (* Timer acabou *)
    timer205_F : BOOL;  (* Timer acabou *)
    timer206_F : BOOL;  (* Timer acabou *)
    timer207_F : BOOL;  (* Timer acabou *)
    timer208_F : BOOL;  (* Timer acabou *)
    timer209_F : BOOL;  (* Timer acabou *)
    timer210_F : BOOL;  (* Timer acabou *)
    timer212_F : BOOL;  (* Timer acabou *)
    timer211_F : BOOL;  (* Timer acabou *)
    timer213_F : BOOL;  (* Timer acabou *)
    timer214_F : BOOL;  (* Timer acabou *)
    timer215_F : BOOL;  (* Timer acabou *)
    timer216_F : BOOL;  (* Timer acabou *)
    timer217_F : BOOL;  (* Timer acabou *)
    timer218_F : BOOL;  (* Timer acabou *)
    timer219_F : BOOL;  (* Timer acabou *)
    timer220_F : BOOL;  (* Timer acabou *)
    Timer221_F : BOOL;  (* Timer acabou *)
    timer222_F : BOOL;  (* Timer acabou *)
    timer223_F : BOOL;  (* Timer acabou *)
    timer224_F : BOOL;  (* Timer acabou *)
    timer225_F : BOOL;  (* Timer acabou *)
    timer226_F : BOOL;  (* Timer acabou *)
    timer227_F : BOOL;  (* Timer acabou *)
    timer228_F : BOOL;  (* Timer acabou *)
    timer229_F : BOOL;  (* Timer acabou *)
    timer230_F : BOOL;  (* Timer acabou *)
    timer231_F : BOOL;  (* Timer acabou *)
    ContadorPecasReparav : CTU;
    ContadorPecasReparaVerdes : CTU;
    ContadorPecasReparaCinzas : CTU;
    Conta_Pecas_Total_Azul : INT;  (* Total de peças azuis *)
    Conta_Pecas_Total_Verde : INT;  (* Total de peças verdes *)
    Conta_Pecas_Total_Cinza : INT;  (* Total de peças cinza *)
    ContaTotalFinalAzul : CTU;
    Conta_Pecas_TotalFinal_Azul : INT;
    timer500_F : BOOL;  (* Timer acabou *)
    timer450 : TON;
    Timer399 : TON;
    timer399_F : BOOL;  (* Timer acabou *)
    ContaTotalFinalVerde : CTU;
    ContaTotalFinalCinza : CTU;
    Timer450_F : BOOL;  (* Timer acabou *)
    ContadorPecasRC : CTU;
    ContadorPecas_Recolha_Comum : INT;
    P0 : REAL;  (* Potenciometro 0 *)
    P1 : REAL;  (* Potenciometro 1 *)
    P2 : REAL;  (* Potenciometro 2 *)
    P3 : REAL;  (* Potenciometro 3 *)
    P4 : REAL;  (* Potenciometro 5 *)
    P5 : REAL;
    Manutencao : INT;
    Flag_ModoManut : BOOL;
    Timer300_F : BOOL;  (* Timer acabou *)
    Timer301_F : BOOL;  (* Timer acabou *)
    Timer300 : TON;
    Timer301 : TON;
    ContaSaida : CTU;
    ContaEntrada : CTU;
    Conta_EntradaTapete : INT;  (* Conta quantas peças entradam no tapete da recolha comum *)
    Conta_Total : INT;  (* Preças totais passadas no tapete *)
END_VAR
VAR_EXTERNAL
    Trama : ARRAY[0..3] OF OEN\Modbus\sModbusReq;
    out_Dig : ARRAY[0..130] OF BOOL;
    in_Dig : ARRAY[0..50] OF BOOL;
    in_Analog : ARRAY[0..10] OF WORD;
    out_Analog : ARRAY[0..10] OF WORD;
    Encomenda_Azul : DINT;  (* Numero de peça desta cor por encomenda *)
    Encomenda_Verde : DINT;  (* Numero de peça desta cor por encomenda *)
    Encomenda_Cinza : DINT;  (* Numero de peça desta cor por encomenda *)
    Peca_Boa_Azul : DINT;  (* Contador de peças boas produzidas *)
    Peca_Boa_Verde : DINT;  (* Contador de peças boas produzidas *)
    Peca_Boa_Cinza : DINT;  (* Contador de peças boas produzidas *)
    Peca_Lixo_Azul : DINT;  (* Contador de peças com defeito produzidas *)
    Peca_Lixo_Verde : DINT;  (* Contador de peças com defeito produzidas *)
    Peca_Lixo_Cinza : DINT;  (* Contador de peças com defeito produzidas *)
    Peca_Stock_Azul : DINT;  (* Contador de peças que foram para stock *)
    Peca_Stock_Verde : DINT;  (* Contador de peças que foram para stock *)
    Peca_Stock_Cinza : DINT;  (* Contador de peças que foram para stock *)
    HMI_Emitter : BOOL;
    HMI_R8 : BOOL;
    HMI_R0 : BOOL;
    HMI_R1 : BOOL;
    HMI_R3 : BOOL;
    HMI_R2 : BOOL;
    HMI_R4 : BOOL;
    HMI_R5 : BOOL;
    HMI_Alarme : BOOL;
    HMI_LG_10 : BOOL;
    HMI_LG_11 : BOOL;
    HMI_LG_12 : BOOL;
    HMI_LG_13 : BOOL;
    HMI_LG_14 : BOOL;
    HMI_LG_15 : BOOL;
    HMI_LG_18 : BOOL;
    HMI_LG_19 : BOOL;
    HMI_LY_10 : BOOL;
    HMI_LY_11 : BOOL;
    HMI_LY_12 : BOOL;
    HMI_LY_13 : BOOL;
    HMI_LY_14 : BOOL;
    HMI_LY_15 : BOOL;
    HMI_LY_18 : BOOL;
    HMI_LY_19 : BOOL;
    HMI_LR_10 : BOOL;
    HMI_LR_11 : BOOL;
    HMI_LR_12 : BOOL;
    HMI_LR_13 : BOOL;
    HMI_LR_14 : BOOL;
    HMI_LR_15 : BOOL;
    HMI_LR_18 : BOOL;
    HMI_LR_19 : BOOL;
    HMI_PP0_X : BOOL;
    HMI_PP1_X : BOOL;
    HMI_PP2_X : BOOL;
    HMI_PP0_Z : BOOL;
    HMI_PP1_Z : BOOL;
    HMI_PP2_Z : BOOL;
    HMI_PP0_Grab : BOOL;
    HMI_PP1_Grab : BOOL;
    HMI_PP2_Grab : BOOL;
    HMI_PP0_CW : BOOL;
    HMI_PP1_CW : BOOL;
    HMI_PP2_CW : BOOL;
    HMI_PP0_CCW : BOOL;
    HMI_PP1_CCW : BOOL;
    HMI_PP2_CCW : BOOL;
    HMI_DS0 : BOOL;
    HMI_DS1 : BOOL;
    HMI_DS2 : BOOL;
    HMI_DS3 : BOOL;
    HMI_DS4 : BOOL;
    HMI_DS5 : BOOL;
    HMI_DS6 : BOOL;
    HMI_DS7 : BOOL;
    HMI_DS8 : BOOL;
    HMI_DS9 : BOOL;
    HMI_DS10 : BOOL;
    HMI_DS11 : BOOL;
    HMI_DS12 : BOOL;
    HMI_DS13 : BOOL;
    HMI_DS14 : BOOL;
    HMI_DS15 : BOOL;
    HMI_DS16 : BOOL;
    HMI_DS17 : BOOL;
    HMI_DS18 : BOOL;
    HMI_DS19 : BOOL;
    HMI_DS20 : BOOL;
    HMI_DS21 : BOOL;
    HMI_DS22 : BOOL;
    HMI_DS23 : BOOL;
    HMI_DS24 : BOOL;
    HMI_DS25 : BOOL;
    HMI_DS26 : BOOL;
    HMI_DS27 : BOOL;
    HMI_DS28 : BOOL;
    HMI_T20 : BOOL;
    HMI_T21 : BOOL;
    HMI_T22 : BOOL;
    HMI_T23 : BOOL;
    HMI_T24 : BOOL;
    HMI_T25 : BOOL;
    HMI_T26 : BOOL;
    HMI_T27 : BOOL;
    HMI_T28 : BOOL;
    HMI_T29 : BOOL;
    HMI_T210 : BOOL;
    HMI_T211 : BOOL;
    HMI_T212 : BOOL;
    HMI_T213 : BOOL;
    HMI_T214 : BOOL;
    HMI_T215 : BOOL;
    HMI_T216 : BOOL;
    HMI_T217 : BOOL;
    HMI_T218 : BOOL;
    HMI_T219 : BOOL;
    HMI_T220 : BOOL;
    HMI_T221 : BOOL;
    HMI_T222 : BOOL;
    HMI_T223 : BOOL;
    HMI_T224 : BOOL;
    HMI_T225 : BOOL;
    HMI_T226 : BOOL;
    HMI_T227 : BOOL;
    HMI_T229 : BOOL;
    HMI_T230 : BOOL;
    HMI_T40 : BOOL;
    HMI_T41 : BOOL;
    HMI_T42 : BOOL;
    HMI_T43 : BOOL;
    HMI_T45 : BOOL;
    HMI_T46 : BOOL;
    HMI_T60 : BOOL;
    HMI_T61 : BOOL;
    HMI_T62 : BOOL;
    HMI_T63 : BOOL;
    HMI_T64 : BOOL;
    HMI_T65 : BOOL;
    HMI_T66 : BOOL;
    HMI_T67 : BOOL;
    HMI_T68 : BOOL;
    HMI_T69 : BOOL;
    HMI_CCW1 : BOOL;
    HMI_CCW0 : BOOL;
    HMI_CW2 : BOOL;
    HMI_CW3 : BOOL;
    HMI_CW4 : BOOL;
    HMI_CW5 : BOOL;
    HMI_CCW6 : BOOL;
    HMI_CCW7 : BOOL;
    HMI_CW8 : BOOL;
    HMI_CW9 : BOOL;
    HMI_CW10 : BOOL;
    HMI_CW11 : BOOL;
    HMI_CW12 : BOOL;
    HMI_CCW14 : BOOL;
    HMI_CW15 : BOOL;
    HMI_CW16 : BOOL;
    HMI_CW17 : BOOL;
    HMI_CW18 : BOOL;
    HMI_CCW20 : BOOL;
    HMI_CW21 : BOOL;
    HMI_PA3_Turn : BOOL;
    HMI_PA4_Turn : BOOL;
    HMI_PA3_Power : BOOL;
    HMI_PA4_Power : BOOL;
    HMI_B0_Power : BOOL;
    HMI_B1_Power : BOOL;
    HMI_B2_Power : BOOL;
    HMI_L0 : BOOL;
    HMI_L1 : BOOL;
    HMI_L2 : BOOL;
    HMI_MCS_0 : BOOL;
    HMI_MCS_1 : BOOL;
    HMI_MCS_2 : BOOL;
    Terminar_sessao : BOOL;
    HMI_BT_Linha_Principal : BOOL;
    HMI_BT_Linha_Azul : BOOL;
    HMI_BT_Linha_Verde : BOOL;
    HMI_BT_Linha_Cinza : BOOL;
    HMI_BT_Linha_Recolha : BOOL;
    Encomenda_Total : DINT;
    HMI_Led_producao : BOOL;
    BTSL_1 : BOOL;  (* Botão Seletor - posição 1 *)
    Page_Access : BOOL;
    Page_Access1 : BOOL;
    HMI_Led_Manutencao : BOOL;
    HMI_VoltaP : BOOL;
    HMI_Volta1 : BOOL;
    HMI_Volta2 : BOOL;
    HMI_Volta3 : BOOL;
    HMI_VoltaRC : BOOL;
    BIO_Input_Bit_00 : BOOL;
    Encomenda_Pronta : BOOL;
    HMI_Flag_Stop : BOOL;
    HMI_VS : DINT;
    HMI_DS29 : BOOL;
    HMI_DS30 : BOOL;
    HMI_DS31 : BOOL;
    HMI_DS33 : BOOL;
    HMI_DS34 : BOOL;
    HMI_DS32 : BOOL;
    BIO_Output_Bit_00 : BOOL;
    BIO_Output_Bit_01 : BOOL;
    BIO_Output_Bit_02 : BOOL;
    ANALOG_Ch1_Analog_Output_Value : INT;
    HMI_Emergencia : BOOL;
END_VAR
VAR
    _e1 : R_TRIG;
    _e2 : R_TRIG;
    _e3 : R_TRIG;
    _e4 : R_TRIG;
    _e5 : R_TRIG;
    _e6 : R_TRIG;
    _e7 : R_TRIG;
    _e8 : R_TRIG;
    _e9 : R_TRIG;
    _e10 : R_TRIG;
    _e11 : R_TRIG;
    _e12 : R_TRIG;
    _e13 : R_TRIG;
    _e14 : R_TRIG;
    _e15 : R_TRIG;
    _e16 : R_TRIG;
    _e17 : R_TRIG;
    _e18 : R_TRIG;
    _e19 : R_TRIG;
    _p20 : BOOL;
    _p21 : BOOL;
    _p22 : BOOL;
    _p23 : BOOL;
    _p24 : BOOL;
    _p25 : BOOL;
    _p26 : BOOL;
    _p27 : BOOL;
    _p28 : BOOL;
    _p29 : BOOL;
    _p30 : BOOL;
    _p31 : BOOL;
    _p32 : BOOL;
    _p33 : BOOL;
    _p34 : BOOL;
    _p35 : BOOL;
    _p36 : BOOL;
    _p37 : BOOL;
    _p38 : BOOL;
    _p39 : BOOL;
    _p40 : BOOL;
END_VAR

(* Section ModBus: ladder, written here as Structured Text *)

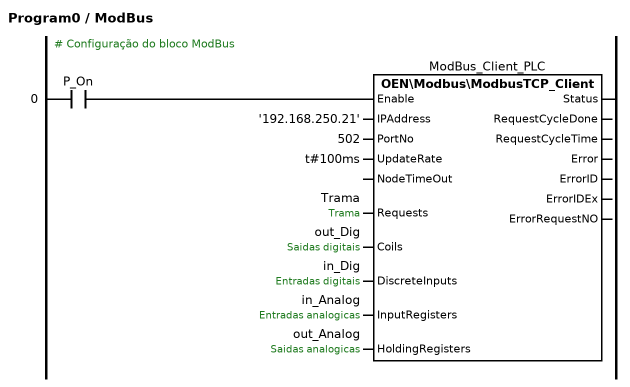
(* Rung 0: # Configuração do bloco ModBus *)
ModBus_Client_PLC(Enable := P_On, IPAddress := '192.168.250.21', PortNo := 502, UpdateRate := t#100ms, Requests := Trama, Coils := out_Dig, DiscreteInputs := in_Dig, InputRegisters := in_Analog, HoldingRegisters := out_Analog);

(* Section Conversoes: ladder, written here as Structured Text *)

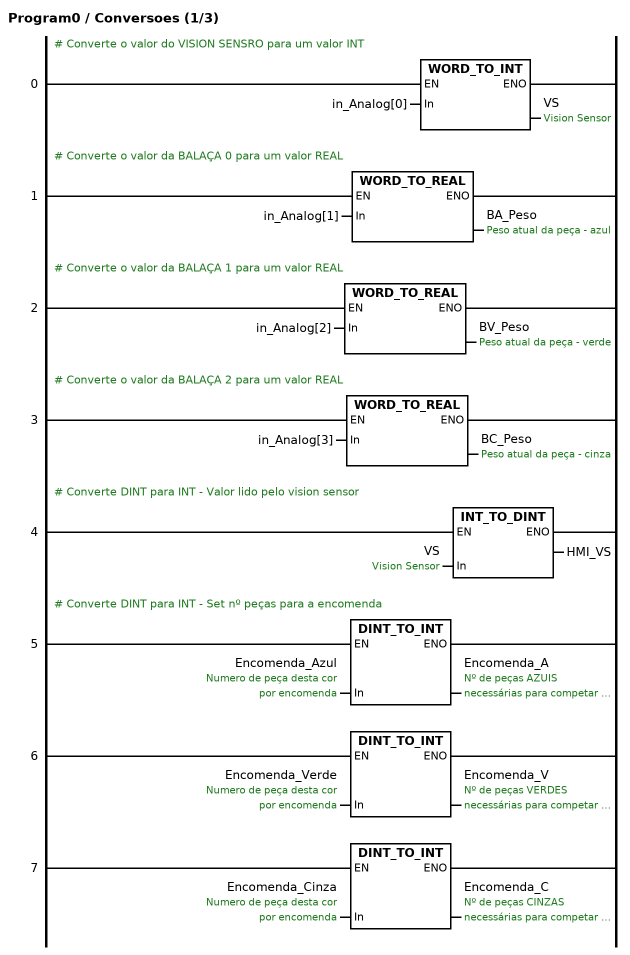
(* Rung 0: # Converte o valor do VISION SENSRO para um valor INT *)
VS := WORD_TO_INT(In := in_Analog[0]);
(* Rung 1: # Converte o valor da BALAÇA 0 para um valor REAL *)
BA_Peso := WORD_TO_REAL(In := in_Analog[1]);
(* Rung 2: # Converte o valor da BALAÇA 1 para um valor REAL *)
BV_Peso := WORD_TO_REAL(In := in_Analog[2]);
(* Rung 3: # Converte o valor da BALAÇA 2 para um valor REAL *)
BC_Peso := WORD_TO_REAL(In := in_Analog[3]);
(* Rung 4: # Converte DINT para INT - Valor lido pelo vision sensor *)
HMI_VS := INT_TO_DINT(In := VS);
(* Rung 5: # Converte DINT para INT - Set nº peças para a encomenda *)
Encomenda_A := DINT_TO_INT(In := Encomenda_Azul);
(* Rung 6 *)
Encomenda_V := DINT_TO_INT(In := Encomenda_Verde);
(* Rung 7 *)
Encomenda_C := DINT_TO_INT(In := Encomenda_Cinza);

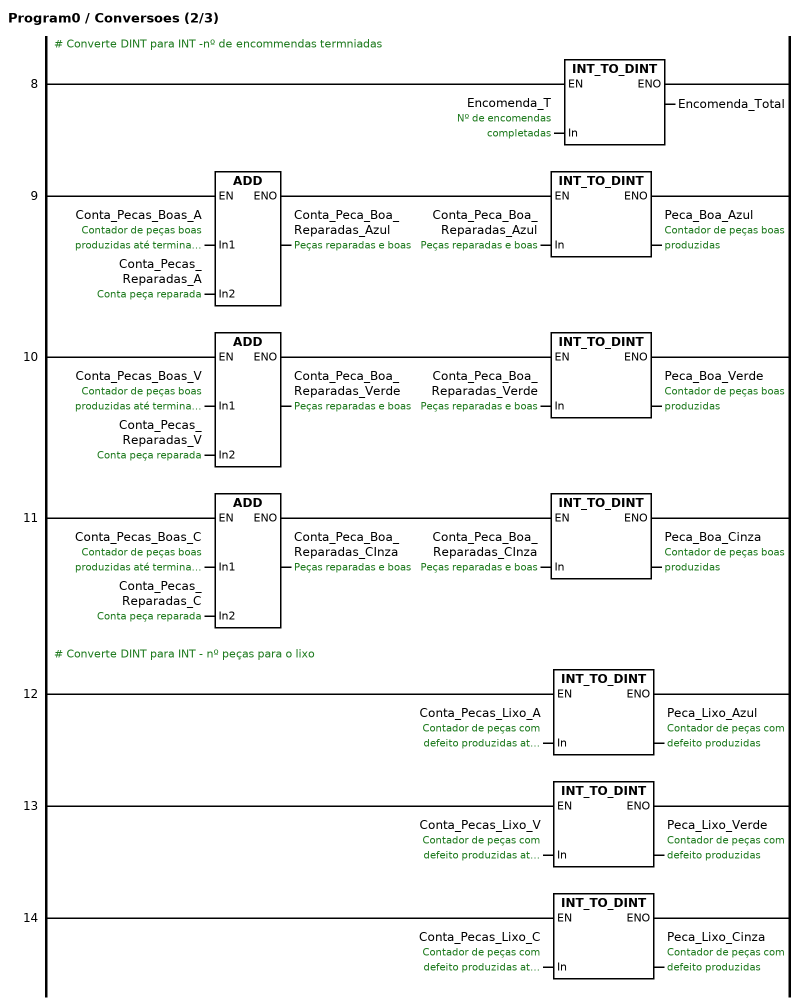
(* Rung 8: # Converte DINT para INT -nº de encommendas termniadas *)
Encomenda_Total := INT_TO_DINT(In := Encomenda_T);
(* Rung 9 *)
Conta_Peca_Boa_Reparadas_Azul := Conta_Pecas_Boas_A + Conta_Pecas_Reparadas_A;
Peca_Boa_Azul := INT_TO_DINT(In := Conta_Peca_Boa_Reparadas_Azul);
(* Rung 10 *)
Conta_Peca_Boa_Reparadas_Verde := Conta_Pecas_Boas_V + Conta_Pecas_Reparadas_V;
Peca_Boa_Verde := INT_TO_DINT(In := Conta_Peca_Boa_Reparadas_Verde);
(* Rung 11 *)
Conta_Peca_Boa_Reparadas_CInza := Conta_Pecas_Boas_C + Conta_Pecas_Reparadas_C;
Peca_Boa_Cinza := INT_TO_DINT(In := Conta_Peca_Boa_Reparadas_CInza);
(* Rung 12: # Converte DINT para INT - nº peças para o lixo *)
Peca_Lixo_Azul := INT_TO_DINT(In := Conta_Pecas_Lixo_A);
(* Rung 13 *)
Peca_Lixo_Verde := INT_TO_DINT(In := Conta_Pecas_Lixo_V);
(* Rung 14 *)
Peca_Lixo_Cinza := INT_TO_DINT(In := Conta_Pecas_Lixo_C);

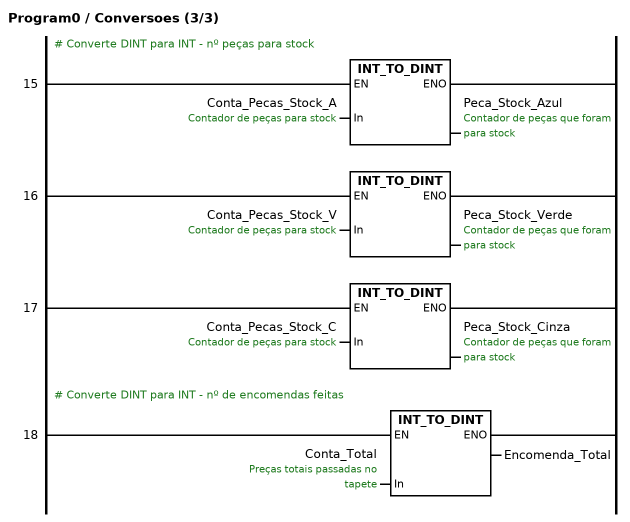
(* Rung 15: # Converte DINT para INT - nº peças para stock *)
Peca_Stock_Azul := INT_TO_DINT(In := Conta_Pecas_Stock_A);
(* Rung 16 *)
Peca_Stock_Verde := INT_TO_DINT(In := Conta_Pecas_Stock_V);
(* Rung 17 *)
Peca_Stock_Cinza := INT_TO_DINT(In := Conta_Pecas_Stock_C);
(* Rung 18: # Converte DINT para INT - nº de encomendas feitas *)
Encomenda_Total := INT_TO_DINT(In := Conta_Total);

(* Section Emergencia: ladder, written here as Structured Text *)

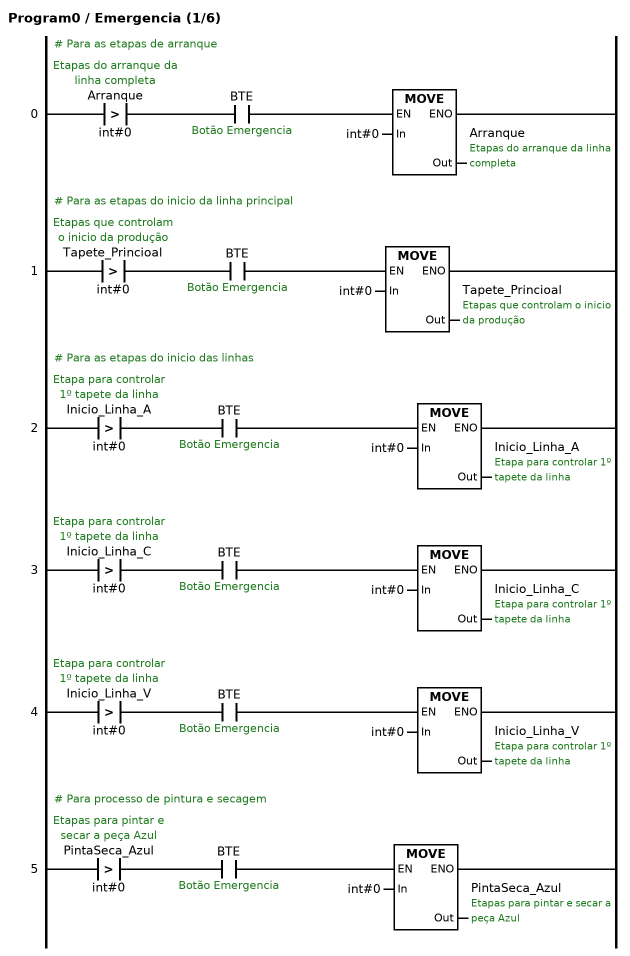
(* Rung 0: # Para as etapas de arranque *)
IF (Arranque > int#0) AND BTE THEN Arranque := int#0; END_IF;
(* Rung 1: # Para as etapas do inicio da linha principal *)
IF (Tapete_Princioal > int#0) AND BTE THEN Tapete_Princioal := int#0; END_IF;
(* Rung 2: # Para as etapas do inicio das linhas *)
IF (Inicio_Linha_A > int#0) AND BTE THEN Inicio_Linha_A := int#0; END_IF;
(* Rung 3 *)
IF (Inicio_Linha_C > int#0) AND BTE THEN Inicio_Linha_C := int#0; END_IF;
(* Rung 4 *)
IF (Inicio_Linha_V > int#0) AND BTE THEN Inicio_Linha_V := int#0; END_IF;
(* Rung 5: # Para processo de pintura e secagem *)
IF (PintaSeca_Azul > int#0) AND BTE THEN PintaSeca_Azul := int#0; END_IF;

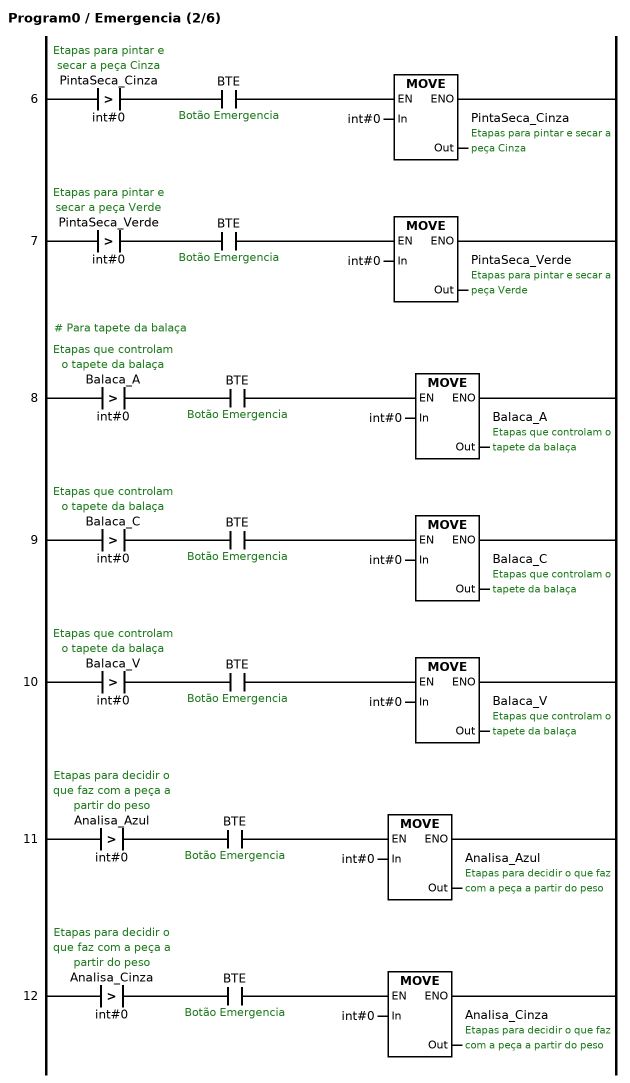
(* Rung 6 *)
IF (PintaSeca_Cinza > int#0) AND BTE THEN PintaSeca_Cinza := int#0; END_IF;
(* Rung 7 *)
IF (PintaSeca_Verde > int#0) AND BTE THEN PintaSeca_Verde := int#0; END_IF;
(* Rung 8: # Para tapete da balaça *)
IF (Balaca_A > int#0) AND BTE THEN Balaca_A := int#0; END_IF;
(* Rung 9 *)
IF (Balaca_C > int#0) AND BTE THEN Balaca_C := int#0; END_IF;
(* Rung 10 *)
IF (Balaca_V > int#0) AND BTE THEN Balaca_V := int#0; END_IF;
(* Rung 11 *)
IF (Analisa_Azul > int#0) AND BTE THEN Analisa_Azul := int#0; END_IF;
(* Rung 12 *)
IF (Analisa_Cinza > int#0) AND BTE THEN Analisa_Cinza := int#0; END_IF;

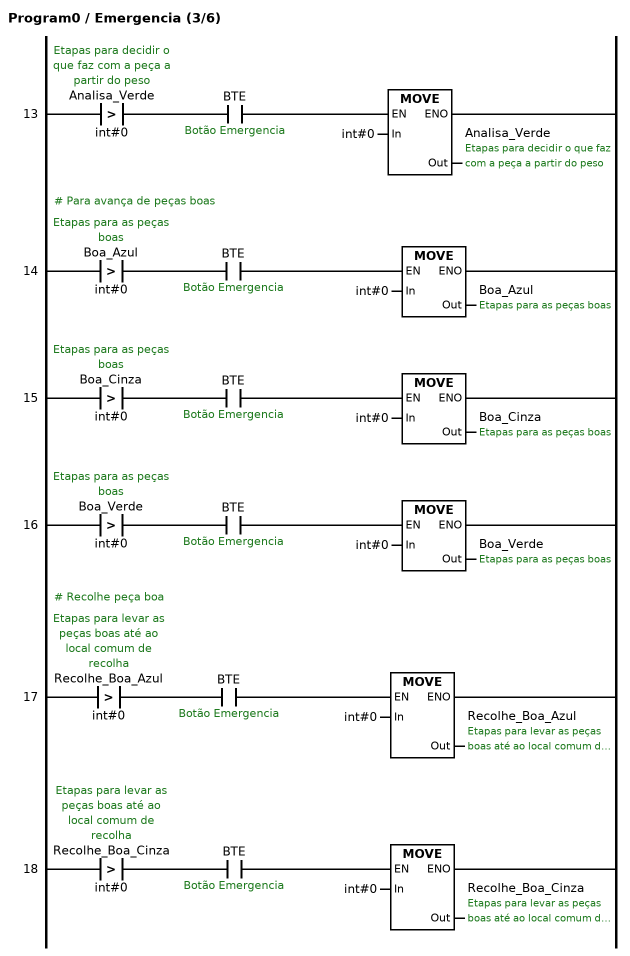
(* Rung 13 *)
IF (Analisa_Verde > int#0) AND BTE THEN Analisa_Verde := int#0; END_IF;
(* Rung 14: # Para avança de peças boas *)
IF (Boa_Azul > int#0) AND BTE THEN Boa_Azul := int#0; END_IF;
(* Rung 15 *)
IF (Boa_Cinza > int#0) AND BTE THEN Boa_Cinza := int#0; END_IF;
(* Rung 16 *)
IF (Boa_Verde > int#0) AND BTE THEN Boa_Verde := int#0; END_IF;
(* Rung 17: # Recolhe peça boa *)
IF (Recolhe_Boa_Azul > int#0) AND BTE THEN Recolhe_Boa_Azul := int#0; END_IF;
(* Rung 18 *)
IF (Recolhe_Boa_Cinza > int#0) AND BTE THEN Recolhe_Boa_Cinza := int#0; END_IF;

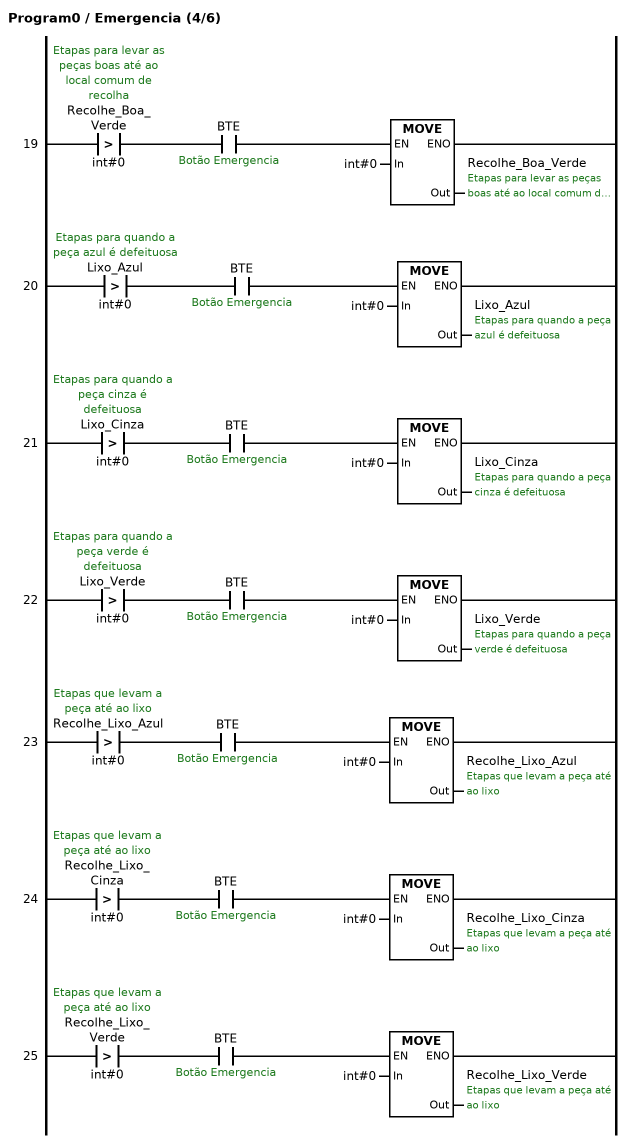
(* Rung 19 *)
IF (Recolhe_Boa_Verde > int#0) AND BTE THEN Recolhe_Boa_Verde := int#0; END_IF;
(* Rung 20 *)
IF (Lixo_Azul > int#0) AND BTE THEN Lixo_Azul := int#0; END_IF;
(* Rung 21 *)
IF (Lixo_Cinza > int#0) AND BTE THEN Lixo_Cinza := int#0; END_IF;
(* Rung 22 *)
IF (Lixo_Verde > int#0) AND BTE THEN Lixo_Verde := int#0; END_IF;
(* Rung 23 *)
IF (Recolhe_Lixo_Azul > int#0) AND BTE THEN Recolhe_Lixo_Azul := int#0; END_IF;
(* Rung 24 *)
IF (Recolhe_Lixo_Cinza > int#0) AND BTE THEN Recolhe_Lixo_Cinza := int#0; END_IF;
(* Rung 25 *)
IF (Recolhe_Lixo_Verde > int#0) AND BTE THEN Recolhe_Lixo_Verde := int#0; END_IF;

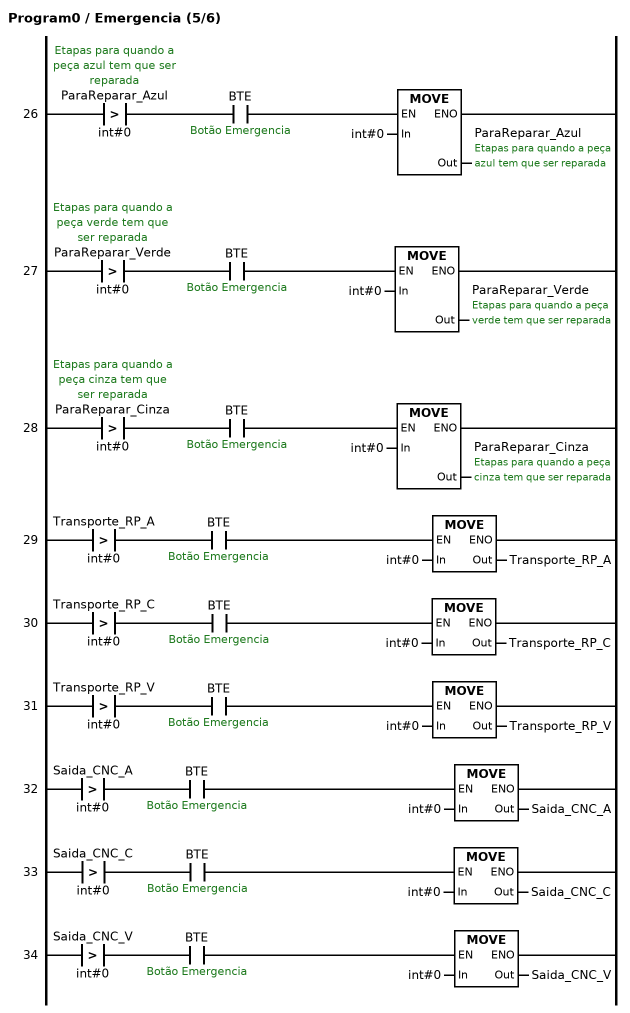
(* Rung 26 *)
IF (ParaReparar_Azul > int#0) AND BTE THEN ParaReparar_Azul := int#0; END_IF;
(* Rung 27 *)
IF (ParaReparar_Verde > int#0) AND BTE THEN ParaReparar_Verde := int#0; END_IF;
(* Rung 28 *)
IF (ParaReparar_Cinza > int#0) AND BTE THEN ParaReparar_Cinza := int#0; END_IF;
(* Rung 29 *)
IF (Transporte_RP_A > int#0) AND BTE THEN Transporte_RP_A := int#0; END_IF;
(* Rung 30 *)
IF (Transporte_RP_C > int#0) AND BTE THEN Transporte_RP_C := int#0; END_IF;
(* Rung 31 *)
IF (Transporte_RP_V > int#0) AND BTE THEN Transporte_RP_V := int#0; END_IF;
(* Rung 32 *)
IF (Saida_CNC_A > int#0) AND BTE THEN Saida_CNC_A := int#0; END_IF;
(* Rung 33 *)
IF (Saida_CNC_C > int#0) AND BTE THEN Saida_CNC_C := int#0; END_IF;
(* Rung 34 *)
IF (Saida_CNC_V > int#0) AND BTE THEN Saida_CNC_V := int#0; END_IF;

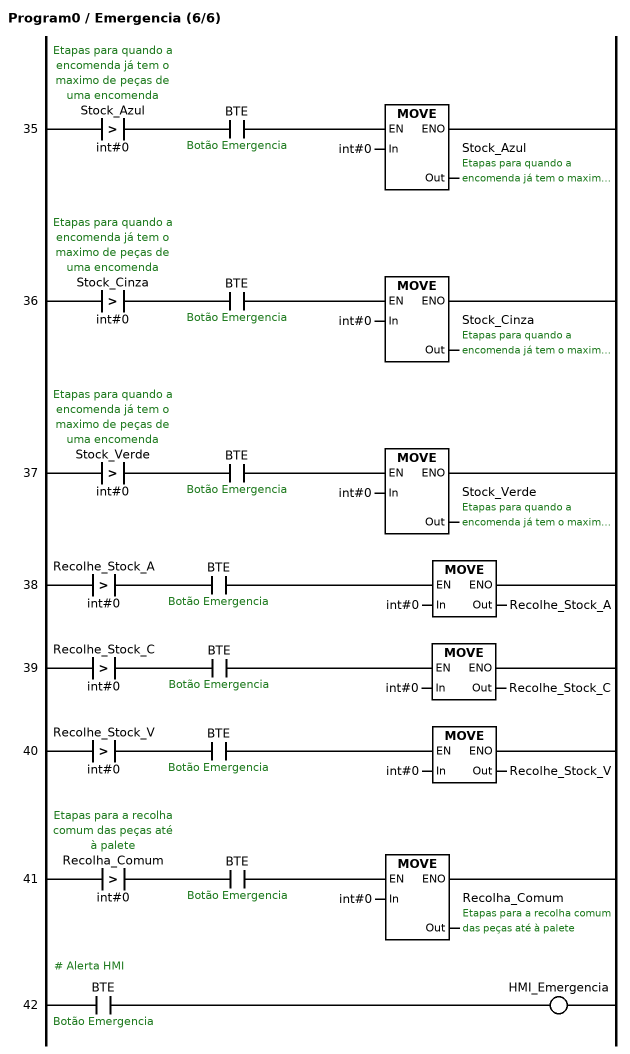
(* Rung 35 *)
IF (Stock_Azul > int#0) AND BTE THEN Stock_Azul := int#0; END_IF;
(* Rung 36 *)
IF (Stock_Cinza > int#0) AND BTE THEN Stock_Cinza := int#0; END_IF;
(* Rung 37 *)
IF (Stock_Verde > int#0) AND BTE THEN Stock_Verde := int#0; END_IF;
(* Rung 38 *)
IF (Recolhe_Stock_A > int#0) AND BTE THEN Recolhe_Stock_A := int#0; END_IF;
(* Rung 39 *)
IF (Recolhe_Stock_C > int#0) AND BTE THEN Recolhe_Stock_C := int#0; END_IF;
(* Rung 40 *)
IF (Recolhe_Stock_V > int#0) AND BTE THEN Recolhe_Stock_V := int#0; END_IF;
(* Rung 41 *)
IF (Recolha_Comum > int#0) AND BTE THEN Recolha_Comum := int#0; END_IF;
(* Rung 42: # Alerta HMI *)
HMI_Emergencia := BTE;

(* Section Contadores: ladder, written here as Structured Text *)

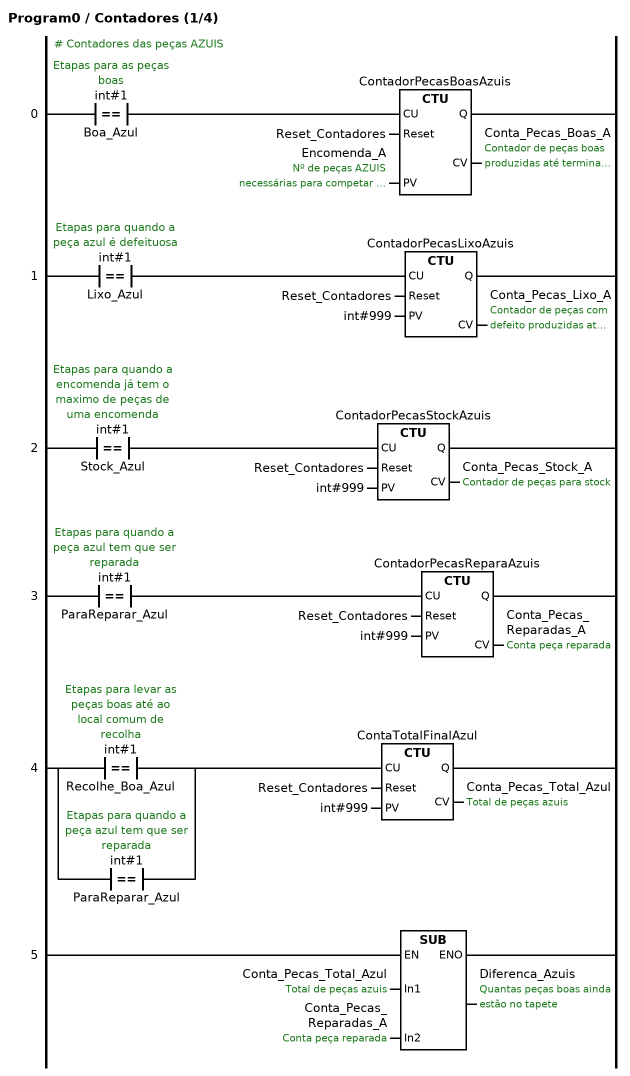
(* Rung 0: # Contadores das peças AZUIS *)
_e1(CLK := int#1 = Boa_Azul);
ContadorPecasBoasAzuis(CU := _e1.Q, Reset := Reset_Contadores, PV := Encomenda_A, CV => Conta_Pecas_Boas_A);
(* Rung 1 *)
_e2(CLK := int#1 = Lixo_Azul);
ContadorPecasLixoAzuis(CU := _e2.Q, Reset := Reset_Contadores, PV := int#999, CV => Conta_Pecas_Lixo_A);
(* Rung 2 *)
_e3(CLK := int#1 = Stock_Azul);
ContadorPecasStockAzuis(CU := _e3.Q, Reset := Reset_Contadores, PV := int#999, CV => Conta_Pecas_Stock_A);
(* Rung 3 *)
_e4(CLK := int#1 = ParaReparar_Azul);
ContadorPecasReparaAzuis(CU := _e4.Q, Reset := Reset_Contadores, PV := int#999, CV => Conta_Pecas_Reparadas_A);
(* Rung 4 *)
_e5(CLK := (int#1 = Recolhe_Boa_Azul) OR (int#1 = ParaReparar_Azul));
ContaTotalFinalAzul(CU := _e5.Q, Reset := Reset_Contadores, PV := int#999, CV => Conta_Pecas_Total_Azul);
(* Rung 5 *)
Diferenca_Azuis := Conta_Pecas_Total_Azul - Conta_Pecas_Reparadas_A;

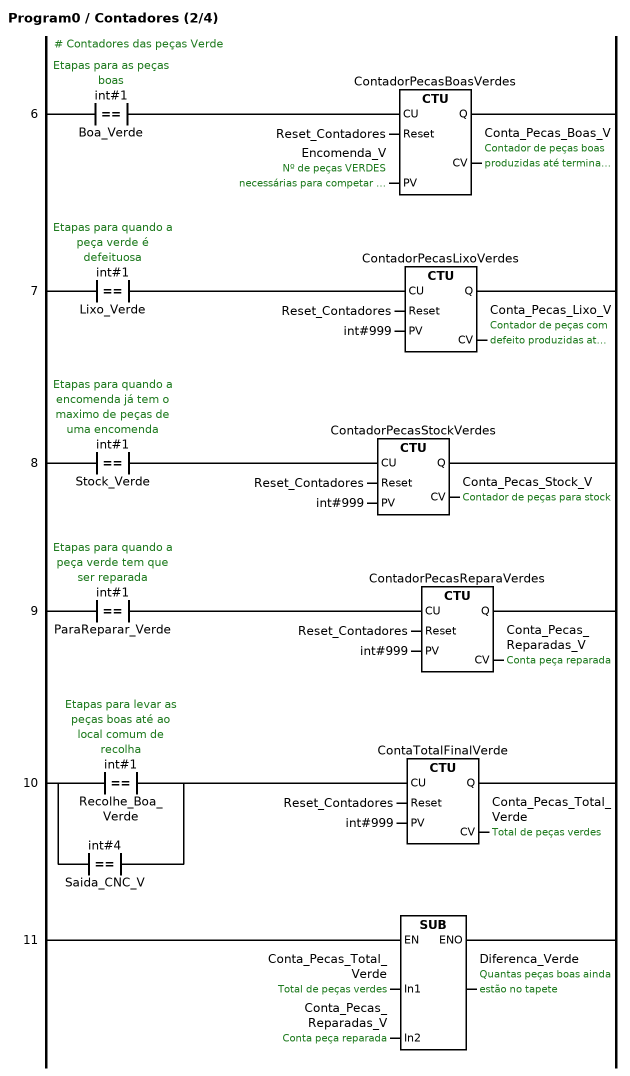
(* Rung 6: # Contadores das peças Verde *)
_e6(CLK := int#1 = Boa_Verde);
ContadorPecasBoasVerdes(CU := _e6.Q, Reset := Reset_Contadores, PV := Encomenda_V, CV => Conta_Pecas_Boas_V);
(* Rung 7 *)
_e7(CLK := int#1 = Lixo_Verde);
ContadorPecasLixoVerdes(CU := _e7.Q, Reset := Reset_Contadores, PV := int#999, CV => Conta_Pecas_Lixo_V);
(* Rung 8 *)
_e8(CLK := int#1 = Stock_Verde);
ContadorPecasStockVerdes(CU := _e8.Q, Reset := Reset_Contadores, PV := int#999, CV => Conta_Pecas_Stock_V);
(* Rung 9 *)
_e9(CLK := int#1 = ParaReparar_Verde);
ContadorPecasReparaVerdes(CU := _e9.Q, Reset := Reset_Contadores, PV := int#999, CV => Conta_Pecas_Reparadas_V);
(* Rung 10 *)
_e10(CLK := (int#1 = Recolhe_Boa_Verde) OR (int#4 = Saida_CNC_V));
ContaTotalFinalVerde(CU := _e10.Q, Reset := Reset_Contadores, PV := int#999, CV => Conta_Pecas_Total_Verde);
(* Rung 11 *)
Diferenca_Verde := Conta_Pecas_Total_Verde - Conta_Pecas_Reparadas_V;

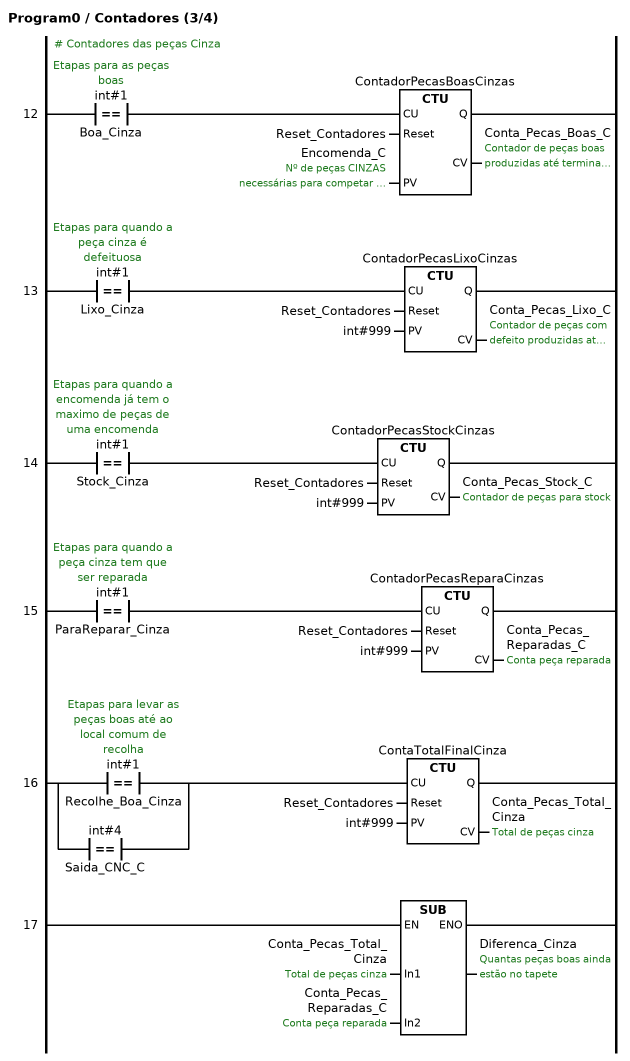
(* Rung 12: # Contadores das peças Cinza *)
_e11(CLK := int#1 = Boa_Cinza);
ContadorPecasBoasCinzas(CU := _e11.Q, Reset := Reset_Contadores, PV := Encomenda_C, CV => Conta_Pecas_Boas_C);
(* Rung 13 *)
_e12(CLK := int#1 = Lixo_Cinza);
ContadorPecasLixoCinzas(CU := _e12.Q, Reset := Reset_Contadores, PV := int#999, CV => Conta_Pecas_Lixo_C);
(* Rung 14 *)
_e13(CLK := int#1 = Stock_Cinza);
ContadorPecasStockCinzas(CU := _e13.Q, Reset := Reset_Contadores, PV := int#999, CV => Conta_Pecas_Stock_C);
(* Rung 15 *)
_e14(CLK := int#1 = ParaReparar_Cinza);
ContadorPecasReparaCinzas(CU := _e14.Q, Reset := Reset_Contadores, PV := int#999, CV => Conta_Pecas_Reparadas_C);
(* Rung 16 *)
_e15(CLK := (int#1 = Recolhe_Boa_Cinza) OR (int#4 = Saida_CNC_C));
ContaTotalFinalCinza(CU := _e15.Q, Reset := Reset_Contadores, PV := int#999, CV => Conta_Pecas_Total_Cinza);
(* Rung 17 *)
Diferenca_Cinza := Conta_Pecas_Total_Cinza - Conta_Pecas_Reparadas_C;

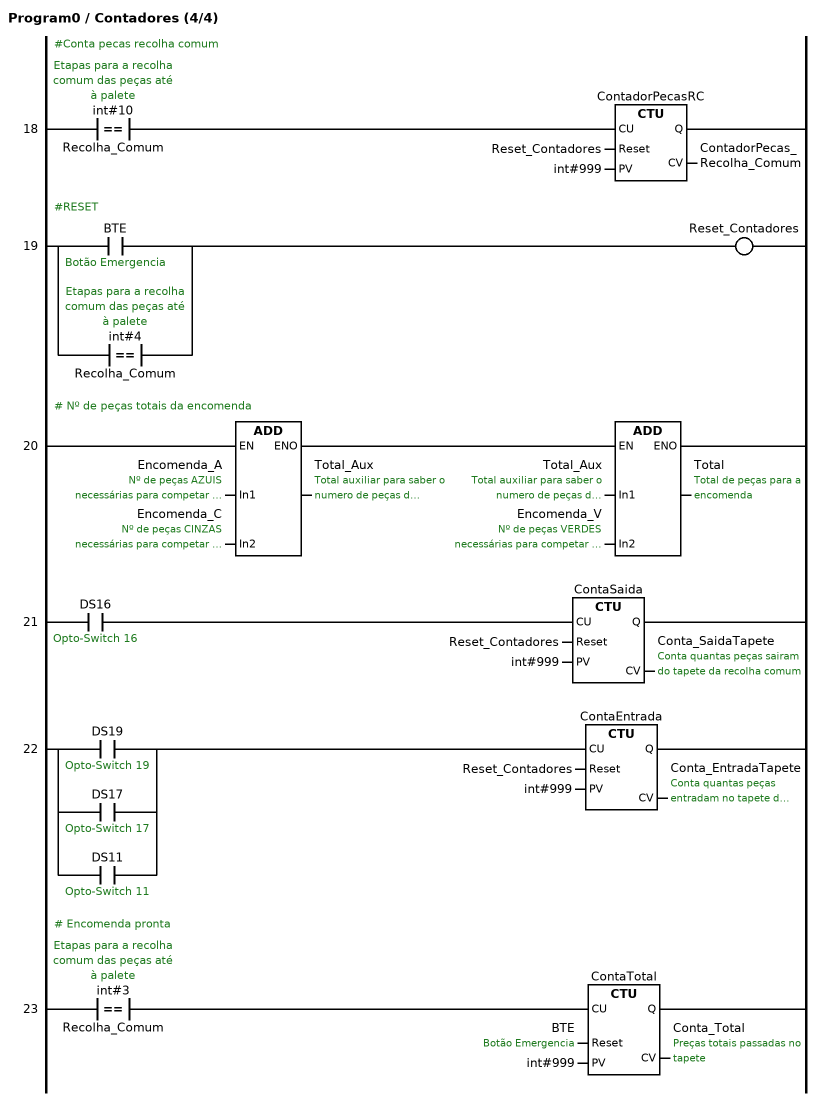
(* Rung 18: #Conta pecas recolha comum *)
_e16(CLK := int#10 = Recolha_Comum);
ContadorPecasRC(CU := _e16.Q, Reset := Reset_Contadores, PV := int#999, CV => ContadorPecas_Recolha_Comum);
(* Rung 19: #RESET *)
Reset_Contadores := BTE OR (int#4 = Recolha_Comum);
(* Rung 20: # Nº de peças totais da encomenda *)
Total_Aux := Encomenda_A + Encomenda_C;
Total := Total_Aux + Encomenda_V;
(* Rung 21 *)
_e17(CLK := DS16);
ContaSaida(CU := _e17.Q, Reset := Reset_Contadores, PV := int#999, CV => Conta_SaidaTapete);
(* Rung 22 *)
_e18(CLK := DS19 OR DS17 OR DS11);
ContaEntrada(CU := _e18.Q, Reset := Reset_Contadores, PV := int#999, CV => Conta_EntradaTapete);
(* Rung 23: # Encomenda pronta *)
_e19(CLK := int#3 = Recolha_Comum);
ContaTotal(CU := _e19.Q, Reset := BTE, PV := int#999, CV => Conta_Total);

(* Section Timeres_Manut: ladder, written here as Structured Text *)

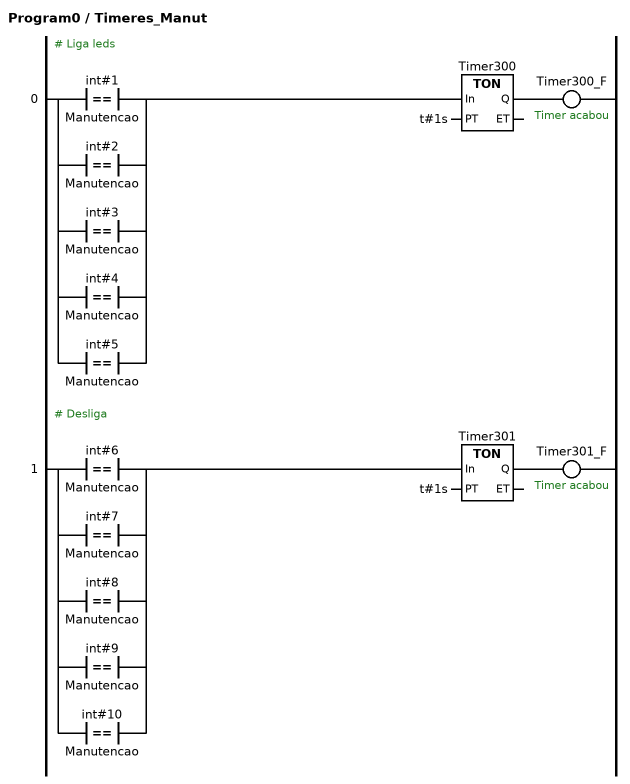
(* Rung 0: # Liga leds *)
Timer300(In := (int#1 = Manutencao) OR (int#2 = Manutencao) OR (int#3 = Manutencao) OR (int#4 = Manutencao) OR (int#5 = Manutencao), PT := t#1s);
Timer300_F := Timer300.Q;
(* Rung 1: # Desliga *)
Timer301(In := (int#6 = Manutencao) OR (int#7 = Manutencao) OR (int#8 = Manutencao) OR (int#9 = Manutencao) OR (int#10 = Manutencao), PT := t#1s);
Timer301_F := Timer301.Q;

(* Section Timeres_Geral: ladder, written here as Structured Text *)

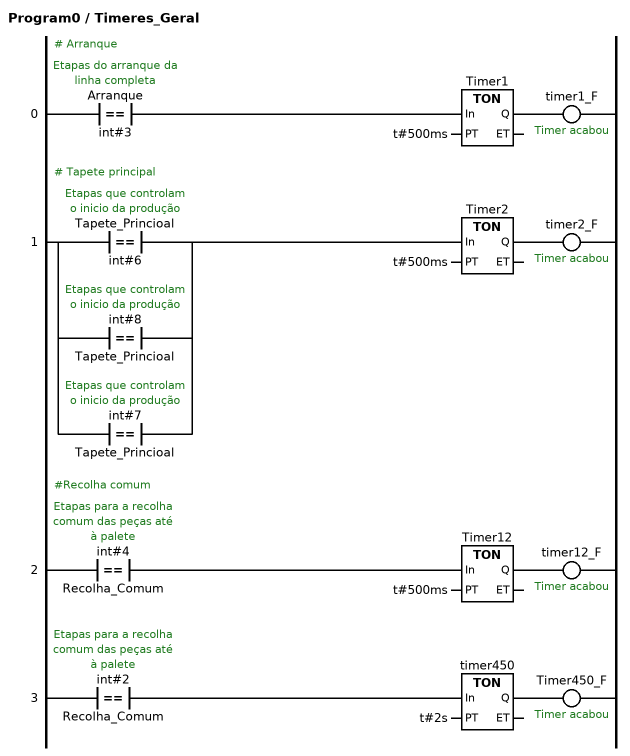
(* Rung 0: # Arranque *)
Timer1(In := Arranque = int#3, PT := t#500ms);
timer1_F := Timer1.Q;
(* Rung 1: # Tapete principal *)
Timer2(In := (Tapete_Princioal = int#6) OR (int#8 = Tapete_Princioal) OR (int#7 = Tapete_Princioal), PT := t#500ms);
timer2_F := Timer2.Q;
(* Rung 2: #Recolha comum *)
Timer12(In := int#4 = Recolha_Comum, PT := t#500ms);
timer12_F := Timer12.Q;
(* Rung 3 *)
timer450(In := int#2 = Recolha_Comum, PT := t#2s);
Timer450_F := timer450.Q;

(* Section Timeres_A: ladder, written here as Structured Text *)

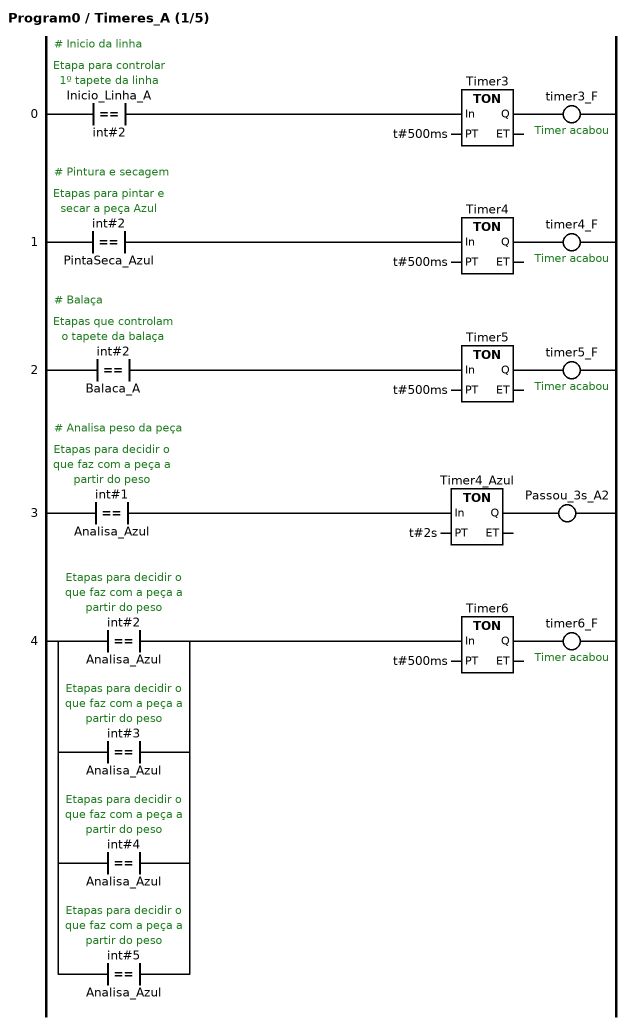
(* Rung 0: # Inicio da linha *)
Timer3(In := Inicio_Linha_A = int#2, PT := t#500ms);
timer3_F := Timer3.Q;
(* Rung 1: # Pintura e secagem *)
Timer4(In := int#2 = PintaSeca_Azul, PT := t#500ms);
timer4_F := Timer4.Q;
(* Rung 2: # Balaça *)
Timer5(In := int#2 = Balaca_A, PT := t#500ms);
timer5_F := Timer5.Q;
(* Rung 3: # Analisa peso da peça *)
Timer4_Azul(In := int#1 = Analisa_Azul, PT := t#2s);
Passou_3s_A2 := Timer4_Azul.Q;
(* Rung 4 *)
Timer6(In := (int#2 = Analisa_Azul) OR (int#3 = Analisa_Azul) OR (int#4 = Analisa_Azul) OR (int#5 = Analisa_Azul), PT := t#500ms);
timer6_F := Timer6.Q;

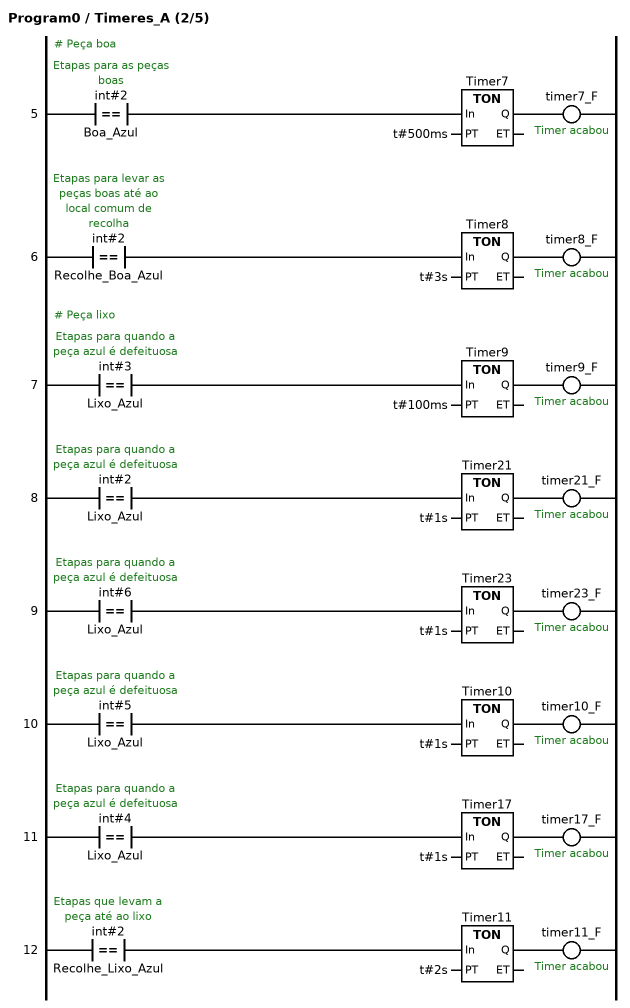
(* Rung 5: # Peça boa *)
Timer7(In := int#2 = Boa_Azul, PT := t#500ms);
timer7_F := Timer7.Q;
(* Rung 6 *)
Timer8(In := int#2 = Recolhe_Boa_Azul, PT := t#3s);
timer8_F := Timer8.Q;
(* Rung 7: # Peça lixo *)
Timer9(In := int#3 = Lixo_Azul, PT := t#100ms);
timer9_F := Timer9.Q;
(* Rung 8 *)
Timer21(In := int#2 = Lixo_Azul, PT := t#1s);
timer21_F := Timer21.Q;
(* Rung 9 *)
Timer23(In := int#6 = Lixo_Azul, PT := t#1s);
timer23_F := Timer23.Q;
(* Rung 10 *)
Timer10(In := int#5 = Lixo_Azul, PT := t#1s);
timer10_F := Timer10.Q;
(* Rung 11 *)
Timer17(In := int#4 = Lixo_Azul, PT := t#1s);
timer17_F := Timer17.Q;
(* Rung 12 *)
Timer11(In := int#2 = Recolhe_Lixo_Azul, PT := t#2s);
timer11_F := Timer11.Q;

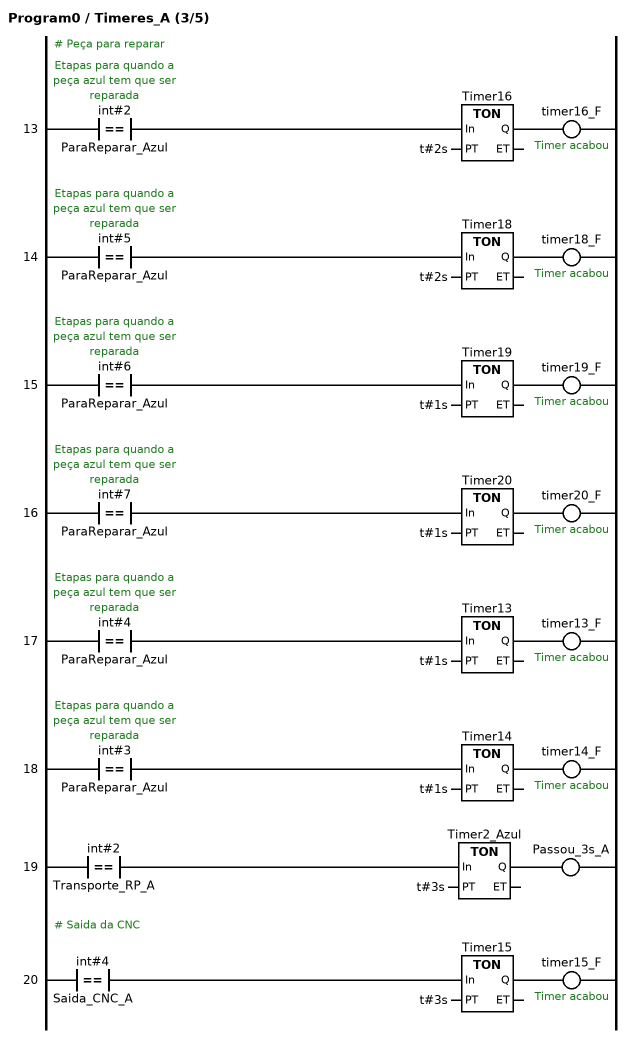
(* Rung 13: # Peça para reparar *)
Timer16(In := int#2 = ParaReparar_Azul, PT := t#2s);
timer16_F := Timer16.Q;
(* Rung 14 *)
Timer18(In := int#5 = ParaReparar_Azul, PT := t#2s);
timer18_F := Timer18.Q;
(* Rung 15 *)
Timer19(In := int#6 = ParaReparar_Azul, PT := t#1s);
timer19_F := Timer19.Q;
(* Rung 16 *)
Timer20(In := int#7 = ParaReparar_Azul, PT := t#1s);
timer20_F := Timer20.Q;
(* Rung 17 *)
Timer13(In := int#4 = ParaReparar_Azul, PT := t#1s);
timer13_F := Timer13.Q;
(* Rung 18 *)
Timer14(In := int#3 = ParaReparar_Azul, PT := t#1s);
timer14_F := Timer14.Q;
(* Rung 19 *)
Timer2_Azul(In := int#2 = Transporte_RP_A, PT := t#3s);
Passou_3s_A := Timer2_Azul.Q;
(* Rung 20: # Saida da CNC *)
Timer15(In := int#4 = Saida_CNC_A, PT := t#3s);
timer15_F := Timer15.Q;

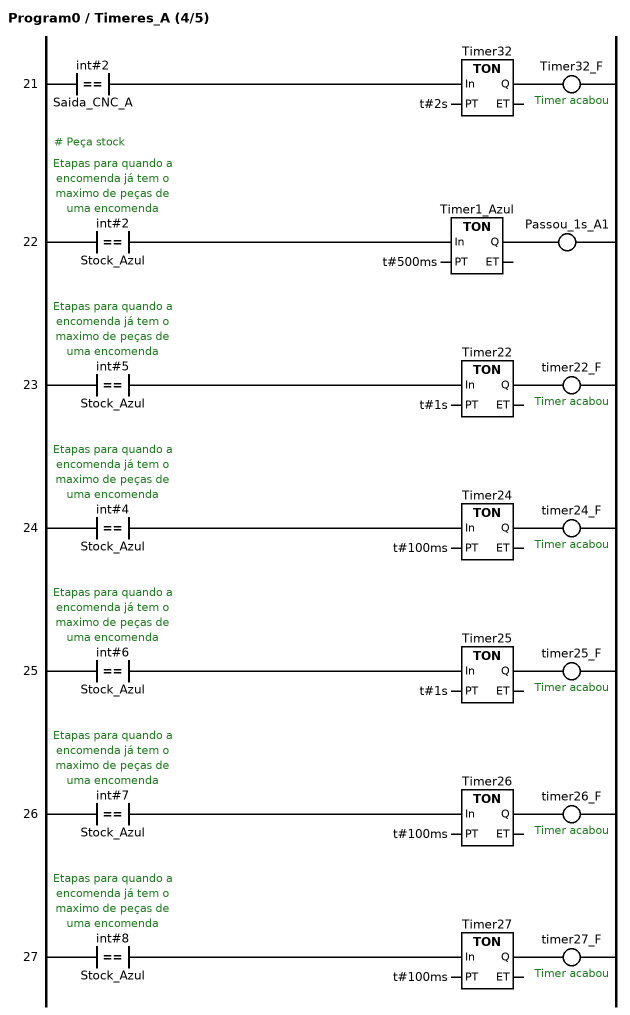
(* Rung 21 *)
Timer32(In := int#2 = Saida_CNC_A, PT := t#2s);
Timer32_F := Timer32.Q;
(* Rung 22: # Peça stock *)
Timer1_Azul(In := int#2 = Stock_Azul, PT := t#500ms);
Passou_1s_A1 := Timer1_Azul.Q;
(* Rung 23 *)
Timer22(In := int#5 = Stock_Azul, PT := t#1s);
timer22_F := Timer22.Q;
(* Rung 24 *)
Timer24(In := int#4 = Stock_Azul, PT := t#100ms);
timer24_F := Timer24.Q;
(* Rung 25 *)
Timer25(In := int#6 = Stock_Azul, PT := t#1s);
timer25_F := Timer25.Q;
(* Rung 26 *)
Timer26(In := int#7 = Stock_Azul, PT := t#100ms);
timer26_F := Timer26.Q;
(* Rung 27 *)
Timer27(In := int#8 = Stock_Azul, PT := t#100ms);
timer27_F := Timer27.Q;

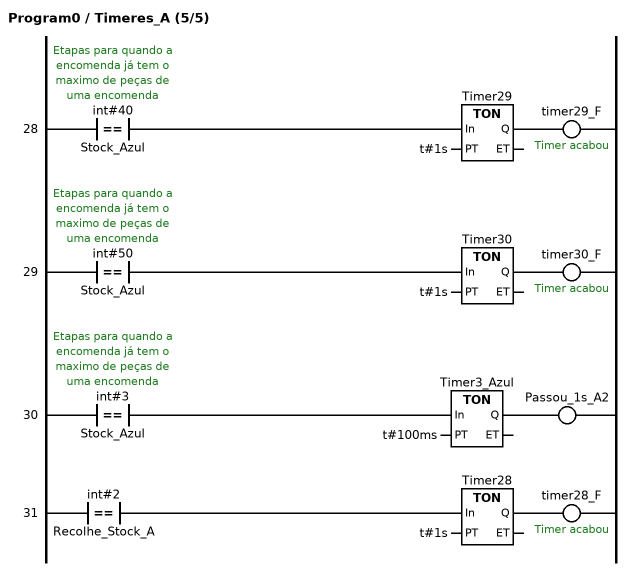
(* Rung 28 *)
Timer29(In := int#40 = Stock_Azul, PT := t#1s);
timer29_F := Timer29.Q;
(* Rung 29 *)
Timer30(In := int#50 = Stock_Azul, PT := t#1s);
timer30_F := Timer30.Q;
(* Rung 30 *)
Timer3_Azul(In := int#3 = Stock_Azul, PT := t#100ms);
Passou_1s_A2 := Timer3_Azul.Q;
(* Rung 31 *)
Timer28(In := int#2 = Recolhe_Stock_A, PT := t#1s);
timer28_F := Timer28.Q;

(* Section Timeres_V: ladder, written here as Structured Text *)

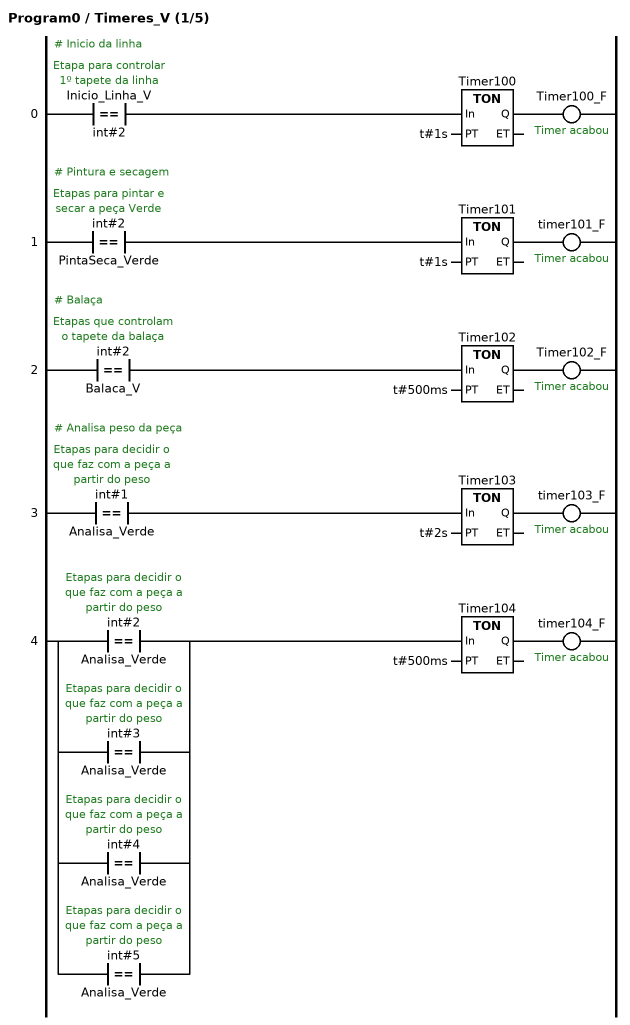
(* Rung 0: # Inicio da linha *)
Timer100(In := Inicio_Linha_V = int#2, PT := t#1s);
Timer100_F := Timer100.Q;
(* Rung 1: # Pintura e secagem *)
Timer101(In := int#2 = PintaSeca_Verde, PT := t#1s);
timer101_F := Timer101.Q;
(* Rung 2: # Balaça *)
Timer102(In := int#2 = Balaca_V, PT := t#500ms);
Timer102_F := Timer102.Q;
(* Rung 3: # Analisa peso da peça *)
Timer103(In := int#1 = Analisa_Verde, PT := t#2s);
timer103_F := Timer103.Q;
(* Rung 4 *)
Timer104(In := (int#2 = Analisa_Verde) OR (int#3 = Analisa_Verde) OR (int#4 = Analisa_Verde) OR (int#5 = Analisa_Verde), PT := t#500ms);
timer104_F := Timer104.Q;

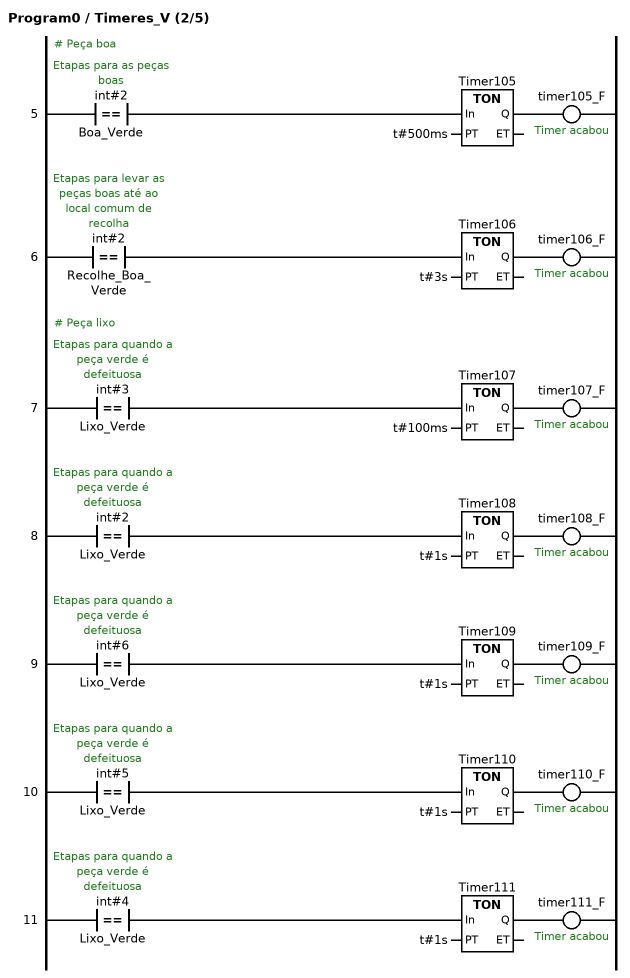
(* Rung 5: # Peça boa *)
Timer105(In := int#2 = Boa_Verde, PT := t#500ms);
timer105_F := Timer105.Q;
(* Rung 6 *)
Timer106(In := int#2 = Recolhe_Boa_Verde, PT := t#3s);
timer106_F := Timer106.Q;
(* Rung 7: # Peça lixo *)
Timer107(In := int#3 = Lixo_Verde, PT := t#100ms);
timer107_F := Timer107.Q;
(* Rung 8 *)
Timer108(In := int#2 = Lixo_Verde, PT := t#1s);
timer108_F := Timer108.Q;
(* Rung 9 *)
Timer109(In := int#6 = Lixo_Verde, PT := t#1s);
timer109_F := Timer109.Q;
(* Rung 10 *)
Timer110(In := int#5 = Lixo_Verde, PT := t#1s);
timer110_F := Timer110.Q;
(* Rung 11 *)
Timer111(In := int#4 = Lixo_Verde, PT := t#1s);
timer111_F := Timer111.Q;

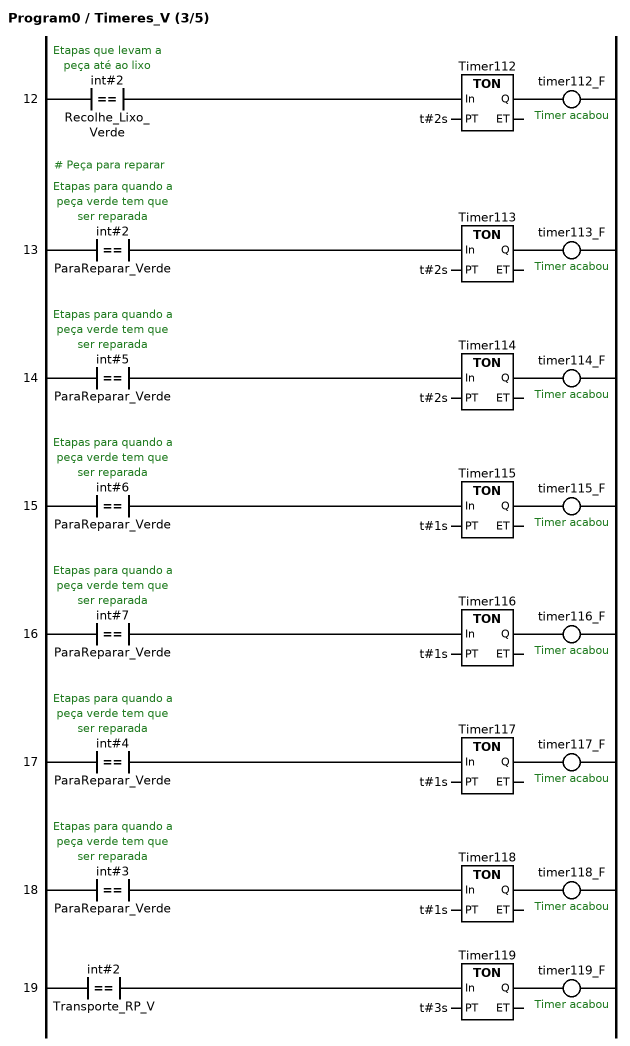
(* Rung 12 *)
Timer112(In := int#2 = Recolhe_Lixo_Verde, PT := t#2s);
timer112_F := Timer112.Q;
(* Rung 13: # Peça para reparar *)
Timer113(In := int#2 = ParaReparar_Verde, PT := t#2s);
timer113_F := Timer113.Q;
(* Rung 14 *)
Timer114(In := int#5 = ParaReparar_Verde, PT := t#2s);
timer114_F := Timer114.Q;
(* Rung 15 *)
Timer115(In := int#6 = ParaReparar_Verde, PT := t#1s);
timer115_F := Timer115.Q;
(* Rung 16 *)
Timer116(In := int#7 = ParaReparar_Verde, PT := t#1s);
timer116_F := Timer116.Q;
(* Rung 17 *)
Timer117(In := int#4 = ParaReparar_Verde, PT := t#1s);
timer117_F := Timer117.Q;
(* Rung 18 *)
Timer118(In := int#3 = ParaReparar_Verde, PT := t#1s);
timer118_F := Timer118.Q;
(* Rung 19 *)
Timer119(In := int#2 = Transporte_RP_V, PT := t#3s);
timer119_F := Timer119.Q;

